(* IEC 61131-3 sources: daoli-st-library/DL_MathData (part 16) *)

(* ---- FC_DL_IntIsPrimeUdint.st ---- *)
(*==============================================================================
 * 组件名称 : FC_DL_IntIsPrimeUdint ｜ 子库 : DL_MathData ｜ v1.0.0 ｜ 2026-11-24
 * 平台     : CODESYS 3.5 / TwinCAT 3 / InoProShop / Machine Expert（纯 IEC，无厂商库）
 * 功能简介 : UDINT 素性判定（试除法）。供伪随机序列、哈希桶数选取、周期分解等调用方。
 *            循环条件写作 nD <= nVal / nD，用除法代替 nD × nD，从根上排除乘法溢出（禁 i*i）。
 * 契约     : 返回 TRUE 表示素数、FALSE 表示合数或 nVal < 2；两者均为合法答案，
 *            bValid := TRUE、bError 保持 FALSE（本件无故障级路径，全为信息级语义）。
 * 依赖     : 无 DL_ 内部依赖（R16 自足实现），无标准库函数调用
 * 错误码   : R297 零码位范式：eErr 恒 0，仅以 bError / bValid 表达
 * 红线自检 : R1 零全局 R2 零%I/%Q R3 纯IEC R4 除零前置（nD ≥ 3 恒定）+ 禁 i*i
 *            R5 双语注释 R6 N/A（无状态机）R7 N/A（无定时器/沿实例）
 *            R10 无类型转换 R11 全声明行分号 R15 标识符零保留字冲突
 * 遗留假设 : nVal < 2（含 0、1）非素数；2 为唯一偶素数，其余偶数短路；
 *            循环天然终止（nD 严格递增、nVal / nD 单调递减），故不设守卫计数；
 *            最坏步数 ⌊√(2³²−1)⌋ / 2 ≈ 32768 次，请在毫秒级任务中避免逐周期调用。
 * 修订历史 : 2026-11-24 R79-B 首版（整数数论族 8/8）
 *============================================================================*)
FUNCTION FC_DL_IntIsPrimeUdint : BOOL
VAR_INPUT
    nVal : UDINT := 0; // 待判定整数 [无量纲] / the value to be tested
END_VAR
VAR_OUTPUT
    eErr   : UDINT; // 错误码，零码位范式恒 0 / error id, always zero under the zero-code rule
    bError : BOOL;  // 故障标志，本件恒 FALSE（素性判定无故障级）/ the fault flag, always FALSE here
    bValid : BOOL;  // 返回值可用标志 / TRUE when the return value is usable
END_VAR
VAR CONSTANT
    DL_ZERO  : UDINT := 0; // 无符号零哨兵 / unsigned zero sentinel
    DL_ONE   : UDINT := 1; // 无符号一哨兵 / unsigned one sentinel
    DL_TWO   : UDINT := 2; // 无符号二哨兵，唯一偶素数 / unsigned two, the only even prime
    DL_THREE : UDINT := 3; // 无符号三哨兵，试除起点 / unsigned three, the trial division start
END_VAR
VAR
    nD : UDINT; // 试除因子，仅取奇数 3, 5, 7, … [无量纲] / the odd trial divisor
END_VAR

// 段 1｜出口预置 / segment 1, preset the exit
FC_DL_IntIsPrimeUdint := FALSE;  // 缺省合数 / default to composite
eErr   := 0;                     // 零码位范式 / zero-code rule
bError := FALSE;                 // 本件无故障级 / this component has no fault level
bValid := FALSE;                 // 判定完成前不认出参 / the result is unusable until the decision is made

// 段 2｜小于 2 的域闸：0 与 1 都不是素数，属合法答案不算故障 / segment 2, the lower domain gate
IF nVal < DL_TWO THEN
    bValid := TRUE;              // FALSE 是合法答案 / FALSE is a legal answer
    RETURN;                      // 返回 FALSE / return the preset FALSE
END_IF

// 段 3｜2 与偶数短路：2 是唯一偶素数 / segment 3, the two and the even number short circuits
IF nVal = DL_TWO THEN
    FC_DL_IntIsPrimeUdint := TRUE;  // 2 为素数 / two is prime
    bValid := TRUE;                 // 判定可用 / the decision is usable
    RETURN;                         // 返回 TRUE / return TRUE
END_IF
IF (nVal MOD DL_TWO) = DL_ZERO THEN
    bValid := TRUE;              // 合数是合法答案 / composite is a legal answer
    RETURN;                      // 返回 FALSE / return the preset FALSE
END_IF

// 段 4｜奇数试除：条件写 nD <= nVal / nD，等价于 nD² <= nVal 但永不溢出 / segment 4, the odd trial division
nD := DL_THREE;                  // 试除起点 3 / start from three
WHILE nD <= (nVal / nD) DO       // 除零不可达：nD ≥ 3 / the divisor is at least three, so no division by zero
    IF (nVal MOD nD) = DL_ZERO THEN
        bValid := TRUE;          // 合数是合法答案 / composite is a legal answer
        RETURN;                  // 返回 FALSE / return the preset FALSE
    END_IF
    nD := nD + DL_TWO;           // 只试奇数 / odd divisors only
END_WHILE

// 段 5｜无因子即素数 / segment 5, no divisor means prime
FC_DL_IntIsPrimeUdint := TRUE;   // 素数 / prime
bValid := TRUE;                  // 判定可用 / the decision is usable
END_FUNCTION

(* ---- FC_DL_IntLcmSafeUdint.st ---- *)
(*==============================================================================
 * 组件名称 : FC_DL_IntLcmSafeUdint ｜ 子库 : DL_MathData ｜ v1.0.0 ｜ 2026-11-24
 * 平台     : CODESYS 3.5 / TwinCAT 3 / InoProShop / Machine Expert（纯 IEC，无厂商库）
 * 功能简介 : UDINT 最小公倍数，先除后乘防溢出：LCM = (nA / GCD) × nB。供脉冲当量配比、
 *            电子齿轮比约分、多轴同步周期归一使用。
 * 契约     : 任一入参为 0 返回 0（IV 约定 LCM(0, x) = 0，信息级，bError 保持 FALSE）；
 *            乘积仍溢出 UDINT 时饱和到 16#FFFF_FFFF 并置 bOverflow := TRUE、bError := TRUE、
 *            bValid := FALSE（饱和值非精确结果，调用方须按故障处理）。
 * 依赖     : 无 DL_ 内部依赖（R16 自足实现：欧几里得 GCD 内联），无标准库函数调用
 * 错误码   : R297 零码位范式：eErr 恒 0，仅以 bError / bValid / bOverflow 表达
 * 红线自检 : R1 零全局 R2 零%I/%Q R3 纯IEC R4 除零前置（nG ≥ 1 由「非双零」保证）+ 乘法前反算上界
 *            R5 双语注释 R6 N/A（无状态机）R7 N/A（无定时器/沿实例）
 *            R10 无类型转换 R11 全声明行分号 R15 标识符零保留字冲突
 * 遗留假设 : 双零入参同属「任一为 0」分支返回 0；GCD 迭代守卫 64 步为安全断言，
 *            理论不可达（欧几里得余量单调递减）；溢出判定用 nQ > (16#FFFF_FFFF / nB)
 *            反算，不做乘法后再比（乘后比已无意义，值已回绕）。
 * 修订历史 : 2026-11-24 R79-B 首版（整数数论族 7/8）
 *============================================================================*)
FUNCTION FC_DL_IntLcmSafeUdint : UDINT
VAR_INPUT
    nA : UDINT := 0; // 左操作数 [脉冲 / 计数] / the left operand, unsigned
    nB : UDINT := 0; // 右操作数 [脉冲 / 计数] / the right operand, unsigned
END_VAR
VAR_OUTPUT
    eErr      : UDINT; // 错误码，零码位范式恒 0 / error id, always zero under the zero-code rule
    bError    : BOOL;  // 乘积溢出时为真（与 bOverflow 同源）/ TRUE on a product overflow, the same source as bOverflow
    bValid    : BOOL;  // 返回值可用标志 / TRUE when the return value is usable
    bOverflow : BOOL;  // 饱和标志：已钳到 16#FFFF_FFFF / TRUE when the result is saturated to the unsigned ceiling
END_VAR
VAR CONSTANT
    DL_ZERO  : UDINT := 0;          // 无符号零哨兵 / unsigned zero sentinel
    DL_ONE   : UDINT := 1;          // 无符号一哨兵 / unsigned one sentinel
    DL_UMAX  : UDINT := 16#FFFF_FFFF; // UDINT 上界，饱和目标 [无量纲] / the unsigned ceiling used for saturation
    DL_GUARD : DINT  := 64;         // GCD 迭代守卫上界 [次] / the euclid guard ceiling
    DL_GUARDI : DINT := 0;          // 迭代计数初值 [次] / the iteration counter start value
END_VAR
VAR
    nX    : UDINT; // GCD 迭代被除数副本 [无量纲] / the gcd dividend copy
    nY    : UDINT; // GCD 迭代除数副本 [无量纲] / the gcd divisor copy
    nG    : UDINT; // 最大公约数 [无量纲] / the greatest common divisor
    nQ    : UDINT; // 先除得商 nA / GCD [无量纲] / the quotient of the division done first
    nIter : DINT;  // GCD 迭代计数，供收敛审计 [次] / the euclid iteration count
END_VAR

// 段 1｜出口预置 / segment 1, preset the exit
FC_DL_IntLcmSafeUdint := DL_ZERO;  // 缺省零 / default zero
eErr      := 0;                    // 零码位范式 / zero-code rule
bError    := FALSE;                // 预置无故障 / preset no fault
bValid    := FALSE;                // 域闸前不认返回值 / the return value is unusable until the gates pass
bOverflow := FALSE;                // 预置未饱和 / preset no saturation

// 段 2｜零入参短路：IV 约定 LCM(0, x) = 0，属信息级不算故障 / segment 2, the zero operand short circuit
IF (nA = DL_ZERO) OR (nB = DL_ZERO) THEN
    bValid := TRUE;                // 0 是合法约定值 / zero is the agreed value here
    RETURN;                        // 返回 0 / return the preset zero
END_IF

// 段 3｜欧几里得 GCD（守卫计数为安全断言，理论不可达）/ segment 3, the euclidean gcd with a guard
nX    := nA;                       // 被除数副本 / dividend copy
nY    := nB;                       // 除数副本 / divisor copy
nIter := DL_GUARDI;                // 计数清零 / clear the counter
WHILE (nY <> DL_ZERO) AND (nIter < DL_GUARD) DO
    nG    := nX MOD nY;            // 余数（nY 非零已证，除法安全）/ the remainder, the divisor is proven non zero
    nX    := nY;                   // 左移 / shift left
    nY    := nG;                   // 左移 / shift left
    nIter := nIter + 1;            // 计数递增 / increment the counter
END_WHILE
IF nIter >= DL_GUARD THEN
    bError := TRUE;                // 守卫命中属平台异常 / a guard hit means a platform anomaly
    RETURN;                        // 返回 0 / return the preset zero
END_IF
nG := nX;                          // 收敛值即 GCD，非双零保证 nG ≥ 1 / the converged value is the gcd and it is at least one

// 段 4｜先除：nQ = nA / GCD，除零已被 nG ≥ 1 拦住 / segment 4, the division done before the multiplication
nQ := nA / nG;                     // 商 [无量纲] / the quotient

// 段 5｜乘法前反算上界：nQ × nB 是否可表示 / segment 5, the pre multiplication ceiling
IF nQ > (DL_UMAX / nB) THEN        // 除零不可达：nB 非零已由段 2 保证 / the divisor is proven non zero
    bOverflow := TRUE;             // 饱和标志 / saturation flag
    bError    := TRUE;             // 故障级：结果不精确 / fault level, the result is inexact
    FC_DL_IntLcmSafeUdint := DL_UMAX;  // 饱和到上界 / saturate to the ceiling
    RETURN;                        // bValid 保持 FALSE / bValid stays FALSE
END_IF

// 段 6｜安全乘法与出口 / segment 6, the safe multiplication and the exit
FC_DL_IntLcmSafeUdint := nQ * nB;  // 已证可表示 / proven representable
bValid := TRUE;                    // 返回值可用 / the return value is usable
END_FUNCTION

(* ---- FC_DL_IntModChk.st ---- *)
(*
    FC_DL_IntModChk —— DINT 整数取模防御包装
    ------------------------------------------------------------------
    组件名称  : FC_DL_IntModChk
    分类      : DL_MathData / IntegerMod
    前缀      : FC_DL_
    版本      : 1.0.0
    溯源      : IEC 61131-3 标准语义的道莅防御性实现（IEC 61131-3 第三版
                整数除法「截断向零」条款 + 余数恒等式 r = a − trunc(a/b)·b
                的防御性落地）；取模语义与判据顺序参照库内 LREAL 域属主
                FC_DL_ModLrealSafe 的闸序（库内复用口径），实现 / 引脚名 /
                码位 100% 自有；clean-room 声明 —— 零代码行复制，无闭源参考。
    平台      : 纯 IEC 61131-3（LINT 64 位整数 + 标准 MOD / DIV 运算符），
                CODESYS 3.5 / TwinCAT 3 / InoProShop / Machine Expert 通用
    作者      : 道莅代码库 · PLC编程专家（R72 构建轮 · 批 1 · 序号 1）
    ------------------------------------------------------------------
    功能说明  : DINT 整数取模 a MOD b 的防御包装，真实工况：齿轮比约分、
                卷绕圈数余量、分度索引回绕前的余数预判。
                判据链顺序：
                ① 除零闸（b = 0 → 故障级早退，输出 0）——先判后除（红线 2）；
                ② DINT_MIN / −1 溢出面闸：被除数 = −2147483648 且除数 = −1 时
                   商 = +2147483648 超出 DINT 可表域（数学余数恒为 0，但三平台
                   MOD 内部实现可能经「先除后乘」路径内溢），此组合显式拦截出
                   信息级，输出确定值 0（数学事实不受影响）；
                ③ 负操作数语义写死：本件**不直接使用平台 MOD 运算符出结果**，
                   而是把两操作数升位到 LINT（64 位，全 DINT 域无损），按
                   IEC 61131-3「整数除法截断向零」标准条款以
                   r = a − trunc(a / b) × b 恒等式自算余数——结果符号**随被除数**
                   （与 C 系 % 口径一致，IEC MOD 主流口径），绝不依赖平台默认；
                ④ 出口（LINT_TO_DINT 降位前已证 |r| < |b| ≤ 2147483648 且
                   r ≠ −2147483648，降位无回绕面）。
                升位理由（可表性反算，R63 口径）：DINT_MIN 取绝对值会在 DINT
                域内回绕（|−2147483648| = 2147483648 > DINT_MAX），任何在
                DINT 域内自算绝对值的写法都带隐藏回绕面；LINT 域内
                ±2147483648 完全可表，升位后全部中间量无回绕。
    错误码    : 16#0002_3900 除数为 0（除零闸命中，输出 0）—— 故障级
                16#0002_3901 被除数 = DINT_MIN 且除数 = −1 的溢出面组合，
                            数学余数恒 0，输出确定值 0、bValid = TRUE —— 信息级，
                            不置 bError（R45）
                加码反证句（R90）：3901 场景（DINT_MIN/−1 组合）无法由「除零码 +
                正常返回值」组合观测——除零码下输出同为 0 但 bValid = FALSE 且
                语义是「除不了」，3901 语义是「可除但实现面危险」，输出组合不可
                互换观测，故立独立码。
    码位总账  : 16#0002_3900 用 ｜ 16#0002_3901 用
    状态机    : N/A —— 纯函数无状态，无 CASE 可写，非法状态不可能出现
    边界与披露: 一 无定时器 / 无沿检测实例 / 无数组下标，周期安全规则 N/A；
                二 零全局变量、零 VAR_EXTERNAL、零物理地址；
                三 整数进位点（终审两式 #2）验收向量：「除子恰为 0」→ 3900
                   故障级输出 0；「被除数 = DINT_MIN 且除子 = −1」→ 3901
                   信息级输出 0；负操作数四象限向量见验收段；
                四 除法面唯一（LINT 域 trunc(a/b)），除数已在段 3 闸为非零，
                   先判后除，无裸除法暴露；
                五 与 FC_DL_ModLrealSafe（DL_MathData，LREAL 浮点域）分工互引：
                   本件只做 DINT 整数域（DINT_MIN/−1 溢出面为浮点域不存在的
                   独立语义），浮点取模一律走属主件，本件不接 LREAL；
                六 依赖声明：仅 Standard.library（无内建函数依赖，LINT 运算符
                   与 DINT_TO_LINT / LINT_TO_DINT 标准转换），三平台无编译门槛。
    验收向量  : V1 (17, 5) → 2；V2 (−17, 5) → −2（符号随被除数）；
                V3 (17, −5) → 2；V4 (−17, −5) → −2；
                V5 (−2147483648, 5) → −3；V6 (−2147483648, −1) → 0 + 3901；
                V7 (x, 0) → 0 + 3900 故障级；V8 (0, 7) → 0。
                算法已证（脚本）：未跑 ｜ 编译器已证（三平台）：未跑
    修订记录  : 2026-11-23 v1.0.0 首次入库（R72 构建轮 · 批 1 · 序号 1）
*)
FUNCTION FC_DL_IntModChk : DINT
VAR_INPUT
    nDividend : DINT;                      (* 被除数，[无量纲整数域] / the dividend, dimensionless integer *)
    nDivisor  : DINT;                      (* 除数，[无量纲整数域]，禁 0 / the divisor, must not be zero *)
END_VAR
VAR_OUTPUT
    bValid    : BOOL;                      (* 返回值（余数）可用标志，故障级为 FALSE / the remainder usable flag, FALSE on fault *)
    bError    : BOOL;                      (* 故障标志，仅故障级码置位（R45 配对）/ the fault flag, raised only on fault level codes *)
    nInfoCode : UDINT;                     (* 信息 / 错误码，0 = 正常 / the info or error id, 0 = ok *)
END_VAR
VAR CONSTANT
    DL_IMD_ZERO   : DINT := 0;             (* 整数零哨兵，除零闸用 [无量纲] / the integer zero sentinel for the divide gate *)
    DL_IMD_DMIN   : DINT := -2147483648;   (* DINT 下界常量（-2^31），溢出面闸用 [无量纲] / the DINT lower bound constant for the overflow gate *)
    DL_IMD_MONE   : DINT := -1;            (* 溢出面除数哨兵 −1 [无量纲] / the overflow gate divisor sentinel *)
END_VAR
VAR
    nLA      : LINT;                       (* 升位被除数（全 DINT 域无损）[无量纲] / the widened dividend *)
    nLB      : LINT;                       (* 升位除数 [无量纲] / the widened divisor *)
    nLQ      : LINT;                       (* LINT 域截断向零商（中间量）[无量纲] / the widened truncating quotient *)
    nLR      : LINT;                       (* LINT 域余数恒等式结果 [无量纲] / the widened remainder *)
END_VAR

// 段 1｜返回值与状态预置（统一出口预置，R256）/ segment 1, preset the return and the status
FC_DL_IntModChk := 0;                      // 故障缺省返回零余数 / the fault default is zero remainder
bValid    := FALSE;                        // 预置不可用，过闸后置位 / preset unusable, set TRUE after the gates
bError    := FALSE;                        // 预置无故障 / preset no fault
nInfoCode := 0;                            // 预置无错 / preset no error
nLA := 0;                                  // 升位中间量清零 / clear the widened dividend
nLB := 0;                                  // 升位中间量清零 / clear the widened divisor
nLQ := 0;                                  // 商中间量清零 / clear the quotient temporary
nLR := 0;                                  // 余数中间量清零 / clear the remainder temporary

// 段 2｜除零闸（先判后除，红线 2；除子恰为 0 验收向量在此命中）/ segment 2, the divide by zero gate
IF nDivisor = DL_IMD_ZERO THEN             // 除数为 0，取模无定义 / the divisor is zero, modulo undefined
    nInfoCode := 16#0002_3900;             // 故障级：除零 / fault level: divide by zero
    bError := TRUE;                        // R45 配对置故障标志 / paired with the fault flag
    bValid := FALSE;                       // 返回值不可用 / the return unusable
    FC_DL_IntModChk := 0;                  // 确定值零出口 / a deterministic zero outlet
    RETURN;                                // 结构早退 / structural exit
END_IF

// 段 3｜DINT_MIN / −1 溢出面闸（商 +2147483648 超 DINT 可表域，防御性拦截）/ segment 3, the DINT_MIN over minus one overflow gate
IF (nDividend = DL_IMD_DMIN) AND (nDivisor = DL_IMD_MONE) THEN // 溢出面组合 / the overflow surface pair
    nInfoCode := 16#0002_3901;             // 信息级：溢出面组合拦截（数学余数恒 0）/ info level: the overflow pair intercepted, the remainder is zero
    bError := FALSE;                       // 信息级不置故障（R45 配对纪律）/ info level never raises a fault
    bValid := TRUE;                        // 数学余数恒为 0，值可用 / the mathematical remainder is zero, usable
    FC_DL_IntModChk := 0;                  // 确定值零出口 / a deterministic zero outlet
    RETURN;                                // 结构早退 / exit
END_IF

// 段 4｜升位与余数恒等式（负操作数语义写死：r = a − trunc(a/b)·b，符号随被除数）/ segment 4, widen and apply the remainder identity
nLA := DINT_TO_LINT(nDividend);            // 被除数升位（全 DINT 域无损）/ widen the dividend lossless
nLB := DINT_TO_LINT(nDivisor);             // 除数升位 / widen the divisor
nLQ := nLA / nLB;                          // IEC 整数除法截断向零（除数已过闸非零）/ the IEC truncating division, divisor gated non zero
nLR := nLA - (nLQ * nLB);                  // 余数恒等式（符号随被除数，不依赖平台 MOD 口径）/ the remainder identity, sign follows the dividend

// 段 5｜降位可表性防线（|r| < |b| ≤ 2147483648 且 r ≠ −2147483648，结构性可证）/ segment 5, the narrowing guard
IF (nLR > DINT_TO_LINT(2147483647)) OR (nLR < DINT_TO_LINT(DL_IMD_DMIN)) THEN // 降位越域防御兜底（不可达，R151 收口纪律）/ the narrowing overflow guard, structurally unreachable
    nInfoCode := 16#0002_3900;             // 复用除零故障级（同属「结果不可信」类，R90 反证：不可达无观测需求）/ reuse the fault code, unreachable
    bError := TRUE;                        // R45 配对置故障标志 / paired with the fault flag
    bValid := FALSE;                       // 返回值不可用 / unusable
    FC_DL_IntModChk := 0;                  // 确定值零出口 / a deterministic zero outlet
    RETURN;                                // 结构早退 / exit
END_IF

// 段 6｜正常出口 / segment 6, the normal outlet
FC_DL_IntModChk := LINT_TO_DINT(nLR);      // 降位发布余数（符号随被除数）/ publish the remainder
bValid := TRUE;                            // 结果可用 / the result usable
END_FUNCTION

(* ---- FC_DL_IntModPowUdint.st ---- *)
(*==============================================================================
 * 组件名称 : FC_DL_IntModPowUdint ｜ 子库 : DL_MathData ｜ v1.0.0 ｜ 2026-11-24
 * 平台     : CODESYS 3.5 / TwinCAT 3 / InoProShop / Machine Expert（纯 IEC，无厂商库）
 * 功能简介 : 模幂运算，返回 nBase^nExp MOD nMod。供校验码、伪随机、整数密钥类运算调用方。
 *            防乘溢出：任何一次乘法都拆成 32 步「加倍-加法」，每步先以「nMod − 加数 是否
 *            够减」判进位再即时归约，故累加积与倍增被乘数恒 < nMod，全程不出现回绕。
 * 契约     : nMod = 0 → 返回 0、bError := TRUE（模数缺失，模幂无定义）；
 *            nMod = 1 → 返回 0、bValid := TRUE（任何数模 1 恒 0，非故障）；
 *            其余 → 返回精确结果、bValid := TRUE、bError 保持 FALSE。
 * 依赖     : 无 DL_ 内部依赖（R16 自足实现：快速乘内联），无标准库函数调用
 * 错误码   : R297 零码位范式：eErr 恒 0，仅以 bError / bValid 表达
 * 红线自检 : R1 零全局 R2 零%I/%Q R3 纯IEC R4 除零前置（nMod ≥ 2 后才有 MOD 与除）+ 乘前归约
 *            R5 双语注释 R6 N/A（无状态机）R7 N/A（无定时器/沿实例）
 *            R10 无类型转换 R11 全声明行分号 R15 标识符零保留字冲突
 * 遗留假设 : 指数位宽固定 UDINT 32 位（内层 FOR 0..31 定长）；两路乘法（nRes × nPow 与
 *            nPow × nPow）合并进同一 32 步循环并行累加，指数位为 0 时积 1 算出后丢弃
 *            （换来「一段代码两用、零重复」，代价是每外层位最多 32 步空转）；
 *            末位之后多做一次倍增无害（nDbl 恒 < nMod），故不设位序守卫。
 * 修订历史 : 2026-11-24 R79-B 首版（整数数论族 9/8 补位）
 *============================================================================*)
FUNCTION FC_DL_IntModPowUdint : UDINT
VAR_INPUT
    nBase : UDINT := 0; // 底数 [无量纲] / the base of the power
    nExp  : UDINT := 0; // 指数 [无量纲] / the exponent
    nMod  : UDINT := 0; // 模数，须 ≥ 2 才有意义 [无量纲] / the modulus, meaningful from two upwards
END_VAR
VAR_OUTPUT
    eErr   : UDINT; // 错误码，零码位范式恒 0 / error id, always zero under the zero-code rule
    bError : BOOL;  // 模数为零时为真 / TRUE when the modulus is zero
    bValid : BOOL;  // 返回值可用标志 / TRUE when the return value is usable
END_VAR
VAR CONSTANT
    DL_ZERO : UDINT := 0; // 无符号零哨兵 / unsigned zero sentinel
    DL_ONE  : UDINT := 1; // 无符号一哨兵 / unsigned one sentinel
    DL_TWO  : UDINT := 2; // 无符号二哨兵，右移与奇偶判据 / unsigned two, the halving and parity base
    DL_BIT0 : DINT  := 0;  // 位循环起点 [位] / the bit loop start index
    DL_BITN : DINT  := 31; // 位循环终点，UDINT 位宽减一 [位] / the bit loop end index
END_VAR
VAR
    nRes  : UDINT; // 结果累加量，恒 < nMod [无量纲] / the result accumulator, always below the modulus
    nPow  : UDINT; // 当前幂底，恒 < nMod [无量纲] / the current power base, always below the modulus
    nExpW : UDINT; // 指数工作副本，逐位右移 [无量纲] / the exponent working copy, shifted per bit
    nMr   : UDINT; // 乘法 1 的乘数（结果量）[无量纲] / the multiplier of the first product
    nMq   : UDINT; // 乘法 2 的乘数（幂底自乘）[无量纲] / the multiplier of the squaring product
    nDbl  : UDINT; // 共用的倍增被乘数，恒 < nMod [无量纲] / the shared doubled multiplicand, always below the modulus
    nAdd  : UDINT; // 本步实际加数，位为 0 时取 0 [无量纲] / the addend of this step, zero on a cleared bit
    nAccR : UDINT; // 乘法 1 的积，恒 < nMod [无量纲] / the accumulator of the first product
    nAccQ : UDINT; // 乘法 2 的积，恒 < nMod [无量纲] / the accumulator of the squaring product
    nBit  : DINT;  // 位循环计数 0..31 [位] / the bit loop counter
END_VAR

// 段 1｜出口预置 / segment 1, preset the exit
FC_DL_IntModPowUdint := DL_ZERO;  // 缺省零 / default zero
eErr   := 0;                      // 零码位范式 / zero-code rule
bError := FALSE;                  // 预置无故障 / preset no fault
bValid := FALSE;                  // 域闸前不认返回值 / the return value is unusable until the gates pass

// 段 2｜模数域闸：零模数故障、一模数恒零 / segment 2, the modulus gates
IF nMod = DL_ZERO THEN
    bError := TRUE;               // 模数缺失，模幂无定义 / without a modulus the operation is undefined
    RETURN;                       // 返回 0 / return the preset zero
END_IF
IF nMod = DL_ONE THEN
    bValid := TRUE;               // 任何数模 1 恒 0，属合法结果 / any value modulo one is zero, a legal result
    RETURN;                       // 返回 0 / return the preset zero
END_IF

// 段 3｜初值：nRes = 1、nPow = nBase MOD nMod（nMod ≥ 2 已证，MOD 安全）/ segment 3, the initial values
nRes  := DL_ONE;                  // 乘法单位元 / the multiplicative identity
nPow  := nBase MOD nMod;          // 底数先归约 / reduce the base first
nExpW := nExp;                    // 指数工作副本 / the exponent working copy

// 段 4｜二进制模幂：指数位自低向高，每轮并行算 nRes × nPow 与 nPow × nPow / segment 4, the binary modular power
WHILE nExpW > DL_ZERO DO
    nMr   := nRes;                // 乘法 1 的乘数 / the first multiplier
    nMq   := nPow;                // 乘法 2 的乘数 / the squaring multiplier
    nDbl  := nPow;                // 两路共用被乘数 / the shared multiplicand
    nAccR := DL_ZERO;             // 积 1 清零 / clear the first accumulator
    nAccQ := DL_ZERO;             // 积 2 清零 / clear the second accumulator
    FOR nBit := DL_BIT0 TO DL_BITN DO
        nAdd := DL_ZERO;                                                     // 加数缺省 0（位为 0 即空加）/ default addend, an empty add on a cleared bit
        IF (nMr MOD DL_TWO) = DL_ONE THEN nAdd := nDbl; END_IF               // 位为 1 才置加数 / load the addend on a set bit
        IF nAccR >= (nMod - nAdd) THEN nAccR := nAccR - (nMod - nAdd); ELSE nAccR := nAccR + nAdd; END_IF  // 加后即时归约，永不溢出 / add and reduce at once
        nAdd := DL_ZERO;                                                     // 加数复用前清零 / clear the reused addend
        IF (nMq MOD DL_TWO) = DL_ONE THEN nAdd := nDbl; END_IF               // 平方路的同款取数 / the same pick for the squaring
        IF nAccQ >= (nMod - nAdd) THEN nAccQ := nAccQ - (nMod - nAdd); ELSE nAccQ := nAccQ + nAdd; END_IF  // 平方路累加 / accumulate the squaring
        nMr := nMr / DL_TWO;                                                 // 乘数 1 右移一位 / shift the first multiplier
        nMq := nMq / DL_TWO;                                                 // 乘数 2 右移一位 / shift the second multiplier
        IF nDbl >= (nMod - nDbl) THEN nDbl := nDbl - (nMod - nDbl); ELSE nDbl := nDbl + nDbl; END_IF        // 被乘数倍增 mod nMod / double the multiplicand modulo the modulus
    END_FOR
    IF (nExpW MOD DL_TWO) = DL_ONE THEN nRes := nAccR; END_IF                // 指数位为 1 才采信积 1 / adopt the first product only on a set exponent bit
    nPow  := nAccQ;               // 平方结果无条件生效 / the squaring always takes effect
    nExpW := nExpW / DL_TWO;      // 指数右移一位 / shift the exponent
END_WHILE

// 段 5｜出口 / segment 5, the exit
FC_DL_IntModPowUdint := nRes;     // 回写结果 / publish the result
bValid := TRUE;                   // 返回值可用 / the return value is usable
END_FUNCTION

(* ---- FC_DL_IntNextPrimeUdint.st ---- *)
(*==============================================================================
 * 组件名称 : FC_DL_IntNextPrimeUdint ｜ 子库 : DL_MathData ｜ v1.0.0 ｜ 2026-11-24
 * 平台     : CODESYS 3.5 / TwinCAT 3 / InoProShop / Machine Expert（纯 IEC，无厂商库）
 * 功能简介 : 求「≥ nVal + 1 的最小素数」（严格大于入参）。供哈希桶数取素数、抖动模数
 *            选取、伪随机种子上限归整使用。试除条件写作 nD <= nCand / nD，禁 i*i 防溢出。
 * 契约     : 找到即返回该素数、bValid := TRUE；nVal ≥ 16#FFFF_FFF0（无足够向上空间）
 *            或 2000 步内未找到（防死循环）或推进中将越过 UDINT 上界 → 返回 0、
 *            bError := TRUE、bValid := FALSE。
 * 依赖     : 无 DL_ 内部依赖（R16 自足实现：试除内联），无标准库函数调用
 * 错误码   : R297 零码位范式：eErr 恒 0，仅以 bError / bValid 表达
 * 红线自检 : R1 零全局 R2 零%I/%Q R3 纯IEC R4 除零前置（nD ≥ 2）+ 步数上限 + 加法溢出兜底
 *            R5 双语注释 R6 N/A（无状态机）R7 N/A（无定时器/沿实例）
 *            R10 无类型转换 R11 全声明行分号 R15 标识符零保留字冲突
 * 遗留假设 : nVal = 0 或 1 时起点取 2（2 是 ≥ 2 的最小素数）；候选逐 1 递增（不跳偶），
 *            保证 2000 步覆盖 2000 个连续整数，远大于 2³² 内的最大素数间隙（≈336），
 *            故「步数命中」只可能发生在接近上界处，与上界兜底互为双保险。
 * 修订历史 : 2026-11-24 R79-B 首版（整数数论族补位）
 *============================================================================*)
FUNCTION FC_DL_IntNextPrimeUdint : UDINT
VAR_INPUT
    nVal : UDINT := 0; // 参考值，本件返回严格大于它的最小素数 [无量纲] / the reference value, the result is strictly above it
END_VAR
VAR_OUTPUT
    eErr   : UDINT; // 错误码，零码位范式恒 0 / error id, always zero under the zero-code rule
    bError : BOOL;  // 无解或搜索步数越界时为真 / TRUE when no answer exists or the search budget is exhausted
    bValid : BOOL;  // 返回值可用标志 / TRUE when the return value is usable
END_VAR
VAR CONSTANT
    DL_ZERO  : UDINT := 0;            // 无符号零哨兵 / unsigned zero sentinel
    DL_ONE   : UDINT := 1;            // 无符号一哨兵 / unsigned one sentinel
    DL_TWO   : UDINT := 2;            // 无符号二哨兵，最小素数 / unsigned two, the smallest prime
    DL_THREE : UDINT := 3;            // 无符号三哨兵，试除起点 / unsigned three, the trial division start
    DL_NEAR  : UDINT := 16#FFFF_FFF0; // 上界保护带起点，超过即判无解 / the guard band start near the ceiling
    DL_GUARD : UDINT := 16#FFFF_FFFE; // 推进溢出兜底线 / the increment overflow guard line
    DL_STEP  : DINT  := 2000;         // 候选搜索步数预算 [步] / the candidate search budget
    DL_STEP0 : DINT  := 0;            // 步数计数初值 [步] / the step counter start value
    DL_STEP1 : DINT  := 1;            // 步数计数步长 [步] / the step counter increment
END_VAR
VAR
    nCand  : UDINT; // 当前候选整数 [无量纲] / the current candidate
    nD     : UDINT; // 试除因子，奇数 3, 5, 7, … [无量纲] / the odd trial divisor
    nStep  : DINT;  // 已消耗的候选步数 [步] / the consumed candidate steps
    bPrime : BOOL;  // 当前候选的素性结论 / the primality verdict of the current candidate
    bFound : BOOL;  // 找到标志 / the found flag
END_VAR

// 段 1｜出口预置 / segment 1, preset the exit
FC_DL_IntNextPrimeUdint := DL_ZERO;  // 缺省零哨兵 / default zero sentinel
eErr    := 0;                        // 零码位范式 / zero-code rule
bError  := FALSE;                    // 预置无故障 / preset no fault
bValid  := FALSE;                    // 域闸前不认返回值 / the return value is unusable until the gates pass

// 段 2｜上界域闸：无足够向上空间即判无解 / segment 2, the ceiling gate
IF nVal >= DL_NEAR THEN
    bError := TRUE;                  // 上界保护带内不搜索 / no search inside the guard band
    RETURN;                          // 返回 0 / return the preset zero
END_IF

// 段 3｜起点：严格大于入参，且不低于 2 / segment 3, the start candidate
nCand  := nVal + DL_ONE;             // 严格大于入参 / strictly above the argument
IF nCand < DL_TWO THEN nCand := DL_TWO; END_IF  // 0/1 的最小数答案是 2 / two is the answer for zero and one
nStep  := DL_STEP0;                  // 步数清零 / clear the step counter
bFound := FALSE;                     // 未找到 / nothing found yet

// 段 4｜候选搜索：逐 1 递增，超出预算即停（防死循环）/ segment 4, the candidate search
WHILE (NOT bFound) AND (nStep < DL_STEP) DO
    nStep  := nStep + DL_STEP1;      // 消耗一步 / consume one step
    bPrime := TRUE;                  // 先假定素数 / assume prime first
    IF (nCand > DL_TWO) AND ((nCand MOD DL_TWO) = DL_ZERO) THEN bPrime := FALSE; END_IF  // 大于 2 的偶数必合数 / every even number above two is composite
    IF bPrime AND (nCand > DL_THREE) THEN
        nD := DL_THREE;              // 试除起点 3 / start from three
        WHILE nD <= (nCand / nD) DO  // 等价于 nD² ≤ nCand 但永不溢出 / equivalent to the square test without overflow
            IF (nCand MOD nD) = DL_ZERO THEN
                bPrime := FALSE;     // 找到因子即合数 / a divisor means composite
                EXIT;                // 跳出试除循环 / leave the trial division loop
            END_IF
            nD := nD + DL_TWO;       // 只试奇数 / odd divisors only
        END_WHILE
    END_IF
    IF bPrime THEN
        bFound := TRUE;              // 候选即答案 / the candidate is the answer
    ELSIF nCand >= DL_GUARD THEN
        bError := TRUE;              // 再推进将越过上界 / another step would overflow the ceiling
        bFound := TRUE;              // 以故障方式结束搜索 / end the search as a fault
        nCand  := DL_ZERO;           // 结果置零哨兵 / force the zero sentinel
    ELSE
        nCand := nCand + DL_ONE;     // 推进到下一候选 / advance to the next candidate
    END_IF
END_WHILE

// 段 5｜出口：未找到（预算耗尽）判故障，找到则回写 / segment 5, the exit
IF (NOT bFound) OR bError THEN
    bError := TRUE;                  // 预算耗尽或无解 / the budget ran out or no answer exists
    RETURN;                          // 返回 0 哨兵 / return the zero sentinel
END_IF
FC_DL_IntNextPrimeUdint := nCand;    // 回写素数 / publish the prime
bValid := TRUE;                      // 返回值可用 / the return value is usable
END_FUNCTION

(* ---- FC_DL_IntPowSatUdint.st ---- *)
(*==============================================================================
 * 组件名称 : FC_DL_IntPowSatUdint ｜ 子库 : DL_MathData ｜ v1.0.2 ｜ 2026-11-24
 * 平台     : CODESYS 3.5 / TwinCAT 3 / InoProShop / Machine Expert（纯 IEC，无厂商库）
 * 功能简介 : 无符号整数快速幂（平方求幂），溢出即饱和到 16#FFFF_FFFF 并置 bOverflow。
 *            乘前反算上界：被乘数 > 上限 DIV 乘数 即判溢出，绝不让乘法先回绕。
 * 契约     : 返回 nBase^nExp；nExp = 0 返回 1（含 0^0 口径取 1）；饱和时返回
 *            16#FFFF_FFFF 且 bOverflow := TRUE，bValid 仍为 TRUE（饱和值是确定结论）。
 * 依赖     : 无 DL_ 内部依赖（R16 自足实现），无标准库函数调用
 * 错误码   : R297 零码位范式：eErr 恒 0，饱和以 bOverflow 表达
 * 红线自检 : R1 零全局 R2 零%I/%Q R3 纯IEC R4 乘前反算防溢出、除零前置、循环上限 32 次
 *            R5 双语注释 R6 N/A（无状态机）R7 N/A（无定时器/沿实例）
 *            R10 无类型转换 R11 全声明行分号 R15 标识符零保留字冲突 R18 N/A（无 bReset）
 * 修订历史 : 2026-11-24 R79-A 首版（整数数论族 5/8）
 *============================================================================*)
FUNCTION FC_DL_IntPowSatUdint : UDINT
VAR_INPUT
    nBase       : UDINT;    // 底数，全域 [无量纲] / base over the whole unsigned range
    nExp        : UDINT;    // 指数，全域 [无量纲] / exponent over the whole unsigned range
END_VAR
VAR_OUTPUT
    eErr        : UDINT;    // 错误码，零码位范式恒 0 / error id, always zero under the zero-code rule
    bError      : BOOL;     // 故障标志，本件结构性不置位 / fault flag, never raised by this component
    bValid      : BOOL;     // 结果可用标志，饱和亦为可用结论 / TRUE even when saturated, saturation is a definite verdict
    bOverflow   : BOOL;     // 结果已饱和到 UDINT 上界 / TRUE when the result saturated at the unsigned upper bound
END_VAR
VAR CONSTANT
    DL_MAX_UDINT : UDINT := 16#FFFF_FFFF;   // UDINT 上界，饱和目标值 [无量纲] / unsigned upper bound and saturation target
    DL_TWO       : UDINT := 2;              // 指数折半基数 [无量纲] / exponent halving radix
    DL_ONE       : UDINT := 1;              // 整数一 / integer one
    DL_ZERO      : UDINT := 0;              // 整数零哨兵 / integer zero sentinel
    DL_ITER_MAX  : UDINT := 32;             // 指数最多 32 位，迭代上限 [次] / an exponent has at most thirty two bits [count]
END_VAR
VAR
    nBaseUse    : UDINT;    // 迭代中的底数（含平方） / running base, includes the squaring steps
    nExpUse     : UDINT;    // 迭代中的指数（逐次折半） / running exponent, halved every step
    nRes        : UDINT;    // 结果累乘器 / result accumulator
    nIter       : UDINT;    // 已用迭代次数 / iterations consumed so far
END_VAR

// 段 1｜出口预置 / segment 1, preset the exit
FC_DL_IntPowSatUdint := 0;      // 缺省 0 / default zero
eErr      := 0;                 // 零码位范式 / zero-code rule
bError    := FALSE;             // 本件不产生故障级 / this component raises no fault
bValid    := TRUE;              // 全定义域给出确定结论 / a definite verdict for the whole domain
bOverflow := FALSE;             // 预置未饱和 / preset unsaturated
nRes      := DL_ONE;            // 累乘器初值 1 / accumulator starts at one

// 段 2｜零指数边界：任何底数的 0 次幂为 1 / segment 2, the zero exponent boundary
IF nExp = DL_ZERO THEN
    FC_DL_IntPowSatUdint := DL_ONE;     // 结果为 1 / the result is one
    RETURN;
END_IF

// 段 3｜平方求幂：逐位判断，乘前反算溢出 / segment 3, square and multiply with an overflow reflection
nBaseUse := nBase;                  // 底数工作副本 / working copy of the base
nExpUse  := nExp;                   // 指数工作副本 / working copy of the exponent
nIter    := DL_ZERO;
WHILE (nExpUse > DL_ZERO) AND (nIter < DL_ITER_MAX) DO
    nIter := nIter + DL_ONE;                        // 守卫自增 / advance the guard
    IF (nExpUse MOD DL_TWO) = DL_ONE THEN           // 当前最低位为 1 才乘 / multiply only when the low bit is set
        IF (nBaseUse <> DL_ZERO) AND (nRes > (DL_MAX_UDINT / nBaseUse)) THEN
            nRes      := DL_MAX_UDINT;              // 反算超界，直接饱和 / the reflection overshoots, saturate at once
            bOverflow := TRUE;
        ELSE
            nRes := nRes * nBaseUse;                // 安全乘法 / safe multiplication
        END_IF
    END_IF
    nExpUse := nExpUse / DL_TWO;                    // 指数折半，除数为常量 2 / halve the exponent
    IF nExpUse > DL_ZERO THEN
        IF (nBaseUse <> DL_ZERO) AND (nBaseUse > (DL_MAX_UDINT / nBaseUse)) THEN
            nBaseUse  := DL_MAX_UDINT;              // 平方超界，钳到上限 / the squaring overshoots, clamp to the ceiling
            bOverflow := TRUE;                      // 平方已越界 = 真溢出（v1.0.2 修：v1.0.1 前此处无回执，静默出残值）/ squaring overflowed, raise the receipt (silent residue before v1.0.2)
        ELSE
            nBaseUse := nBaseUse * nBaseUse;        // 安全平方 / safe squaring
        END_IF
    END_IF
END_WHILE
(* v1.0.2 更正：v1.0.1 曾在此按 nIter 触顶置 bOverflow，但 nBase <= 1 且 nExp >= 2^31 时
   循环合法打满 32 次仍应收敛（1^N = 1），该判据造成假溢出回执，已删除；
   溢出回执改为只在「乘前反算越界」与「平方钳位」两处产生（唯一真溢出来源）。 *)

// 段 4｜出口 / segment 4, exit
FC_DL_IntPowSatUdint := nRes;                   // 结果或饱和值 / the result or the saturation value
END_FUNCTION

(* ---- FC_DL_IntReverseDigitsUdint.st ---- *)
(*==============================================================================
 * 组件名称 : FC_DL_IntReverseDigitsUdint ｜ 子库 : DL_MathData ｜ v1.0.0 ｜ 2026-11-24
 * 平台     : CODESYS 3.5 / TwinCAT 3 / InoProShop / Machine Expert（纯 IEC，无厂商库）
 * 功能简介 : 无符号整数的十进制数字反转（如 123 → 321，120 → 21，末尾零自然丢弃）。
 *            逐位取余乘十再累加，纯整数实现。乘前反算：累加器 > (上界 − 当前位) DIV 10
 *            即判溢出，饱和到 16#FFFF_FFFF 并置 bOverflow。
 * 契约     : 返回反转值；反转结果超 UDINT 域时返回 16#FFFF_FFFF、bOverflow := TRUE、
 *            bValid 保持 TRUE（饱和值是确定结论）。nVal = 0 返回 0。
 * 依赖     : 无 DL_ 内部依赖（R16 自足实现），无标准库函数调用
 * 错误码   : R297 零码位范式：eErr 恒 0，溢出以 bOverflow 表达
 * 红线自检 : R1 零全局 R2 零%I/%Q R3 纯IEC R4 乘前反算防溢出、循环上界 10 次、除数为常量
 *            R5 双语注释 R6 N/A（无状态机）R7 N/A（无定时器/沿实例）
 *            R10 无类型转换 R11 全声明行分号 R15 标识符零保留字冲突 R18 N/A（无 bReset）
 * 修订历史 : 2026-11-24 R79-A 首版（整数数论族 8/8）
 *============================================================================*)
FUNCTION FC_DL_IntReverseDigitsUdint : UDINT
VAR_INPUT
    nVal        : UDINT;    // 待反转整数，全域 0~16#FFFF_FFFF [无量纲] / value to reverse over the whole unsigned range
END_VAR
VAR_OUTPUT
    eErr        : UDINT;    // 错误码，零码位范式恒 0 / error id, always zero under the zero-code rule
    bError      : BOOL;     // 故障标志，本件结构性不置位 / fault flag, never raised by this component
    bValid      : BOOL;     // 结果可用标志，饱和亦为可用结论 / TRUE even when saturated
    bOverflow   : BOOL;     // 反转结果已饱和到 UDINT 上界 / TRUE when the reversed value saturated
END_VAR
VAR CONSTANT
    DL_TEN       : UDINT := 10;             // 十进制基数 [无量纲] / decimal radix, dimensionless
    DL_MAX_UDINT : UDINT := 16#FFFF_FFFF;   // UDINT 上界，饱和目标值 [无量纲] / unsigned upper bound and saturation target
    DL_ZERO      : UDINT := 0;              // 整数零哨兵 / integer zero sentinel
    DL_LOOP_MAX  : UDINT := 10;             // UDINT 十进制最大位数，循环上界 [位] / loop cap equal to the largest decimal width [digit]
END_VAR
VAR
    nRest       : UDINT;    // 降位过程中的剩余值 / remaining value while descending
    nRev        : UDINT;    // 反转累加器 / reversed accumulator
    nDigit      : UDINT;    // 当前取出的个位数 / the digit taken from the current position
    nGuard      : UDINT;    // 循环守卫计数 / loop guard counter
END_VAR

// 段 1｜出口预置 / segment 1, preset the exit
FC_DL_IntReverseDigitsUdint := 0;   // 缺省 0 / default zero
eErr      := 0;                     // 零码位范式 / zero-code rule
bError    := FALSE;                 // 本件不产生故障级 / this component raises no fault
bValid    := TRUE;                  // 饱和也是确定结论 / saturation is still a definite verdict
bOverflow := FALSE;                 // 预置未饱和 / preset unsaturated
nRest     := nVal;                  // 从输入起步 / start from the input
nRev      := DL_ZERO;               // 累加器清零 / clear the accumulator
nGuard    := DL_ZERO;               // 守卫清零 / clear the guard

// 段 2｜逐位反转：取个位 → 降位 → 乘前反算后累加 / segment 2, digit by digit reversal with an overflow reflection
WHILE (nRest <> DL_ZERO) AND (nGuard < DL_LOOP_MAX) DO
    nGuard := nGuard + 1;                                   // 守卫自增 / advance the guard
    nDigit := nRest MOD DL_TEN;                             // 取个位 / take the units digit
    nRest  := nRest / DL_TEN;                               // 降一位 / shift one digit down
    IF nRev > ((DL_MAX_UDINT - nDigit) / DL_TEN) THEN
        nRev      := DL_MAX_UDINT;                          // 反算超界，饱和退出 / the reflection overshoots, saturate and stop
        bOverflow := TRUE;
        EXIT;
    END_IF
    nRev := (nRev * DL_TEN) + nDigit;                       // 旧位左移一位并接上新位 / shift the old digits and append
END_WHILE

// 段 3｜出口 / segment 3, exit
FC_DL_IntReverseDigitsUdint := nRev;    // 反转值或饱和值 / the reversed value or the saturation value
END_FUNCTION

(* ---- FC_DL_IntSqrtFloorUdint.st ---- *)
(*==============================================================================
 * 组件名称 : FC_DL_IntSqrtFloorUdint ｜ 子库 : DL_MathData ｜ v1.0.0 ｜ 2026-11-24
 * 平台     : CODESYS 3.5 / TwinCAT 3 / InoProShop / Machine Expert（纯 IEC，无厂商库）
 * 功能简介 : 无符号整数平方根向下取整 ⌊√nVal⌋。牛顿迭代：初值 nVal DIV 2 + 1，
 *            下一试值 = (试值 + nVal DIV 试值) DIV 2，试值不再下降即收敛。
 *            纯整数运算，无浮点、无 SQRT，2^32 全域精确。
 * 契约     : 返回 ⌊√nVal⌋；nVal = 0 返回 0；nIter 达上限 64 次仍未收敛时返回最后一次
 *            试值并置 bError（结构性不可达，作为防死循环兜底）。
 * 依赖     : 无 DL_ 内部依赖（R16 自足实现），无标准库函数调用
 * 错误码   : R297 零码位范式：eErr 恒 0，仅以 bError / bValid 表达
 * 红线自检 : R1 零全局 R2 零%I/%Q R3 纯IEC R4 除零前置（试值恒 ≥1）、迭代上限兜底、
 *            和式上界 ≤ 2^31+1 不溢出 R5 双语注释 R6 N/A（无状态机）
 *            R7 N/A（无定时器/沿实例）R10 无类型转换 R11 全声明行分号
 *            R15 标识符零保留字冲突 R18 N/A（无 bReset）
 * 修订历史 : 2026-11-24 R79-A 首版（整数数论族 1/8）
 *============================================================================*)
FUNCTION FC_DL_IntSqrtFloorUdint : UDINT
VAR_INPUT
    nVal        : UDINT;    // 被开方数，全域 0~16#FFFF_FFFF [无量纲] / radicand over the whole unsigned range
END_VAR
VAR_OUTPUT
    eErr        : UDINT;    // 错误码，零码位范式恒 0 / error id, always zero under the zero-code rule
    bError      : BOOL;     // 迭代未收敛为真（结构性不可达） / TRUE when the iteration fails to converge, unreachable in theory
    bValid      : BOOL;     // 结果可用标志 / result usable flag
END_VAR
VAR CONSTANT
    DL_TWO      : UDINT := 2;               // 牛顿迭代的除数 2 [无量纲] / Newton divisor, dimensionless
    DL_ONE      : UDINT := 1;               // 整数一 [无量纲] / integer one, dimensionless
    DL_ZERO     : UDINT := 0;               // 整数零哨兵 [无量纲] / integer zero sentinel, dimensionless
    DL_ITER_MAX : UDINT := 64;              // 迭代次数上限，二次收敛下 32 次已足 [次] / iteration cap, quadratic convergence needs far fewer [count]
END_VAR
VAR
    nApprox     : UDINT;    // 当前试值，迭代中单调下降 / current trial value, monotonically decreasing
    nNext       : UDINT;    // 下一试值 / next trial value
    nIter       : UDINT;    // 已用迭代次数 / iterations consumed so far
END_VAR

// 段 1｜出口预置 / segment 1, preset the exit
FC_DL_IntSqrtFloorUdint := 0;   // 缺省 0 / default zero
eErr   := 0;                    // 零码位范式 / zero-code rule
bError := FALSE;                // 预置无故障 / preset no fault
bValid := FALSE;                // 计算完成前不认结果 / unusable until the iteration ends

// 段 2｜零边界：0 的平方根为 0，直接放行，避免初值 1 走迭代 / segment 2, the zero boundary
IF nVal = DL_ZERO THEN
    bValid := TRUE;             // 结果 0 可用 / the zero result is usable
    RETURN;                     // 返回 0 / return zero
END_IF

// 段 3｜牛顿迭代：初值取 nVal DIV 2 + 1，必 ≥ √nVal，故单调下降 / segment 3, Newton iteration from an upper bound
nApprox := (nVal / DL_TWO) + DL_ONE;                // 上界初值，避免 nVal DIV nApprox 除零 / upper bound start, keeps the divisor non zero
nIter   := DL_ZERO;                                 // 迭代计数清零 / clear the counter
WHILE nIter < DL_ITER_MAX DO
    nIter   := nIter + DL_ONE;                      // 先计数后算，保证上限生效 / count first so the cap is honoured
    nNext   := (nApprox + (nVal / nApprox)) / DL_TWO;   // 和式上界约 2^31+1，不溢出 / the sum stays near two to the thirty first, no overflow
    IF nNext >= nApprox THEN
        EXIT;                                       // 试值不再下降即收敛 / the trial stops decreasing, converged
    END_IF
    nApprox := nNext;                               // 继续下降 / keep descending
END_WHILE

// 段 4｜收敛自证：用尽上限仍未收敛按故障处置，返回最后一次试值 / segment 4, convergence self proof
IF nIter >= DL_ITER_MAX THEN
    bError := TRUE;                 // 未收敛（理论不可达）/ not converged, unreachable in theory
    FC_DL_IntSqrtFloorUdint := nApprox;
    RETURN;                         // 返回最后一次试值，bValid 保持 FALSE / return the last trial with bValid still FALSE
END_IF

// 段 5｜出口 / segment 5, exit
FC_DL_IntSqrtFloorUdint := nApprox;     // ⌊√nVal⌋ / floor of the square root
bValid := TRUE;                         // 结果可用 / the result is usable
END_FUNCTION

(* ---- FC_DL_IntToFixedField.st ---- *)
(*==============================================================================
 * 组件名称 (Component)  : FC_DL_IntToFixedField
 * 溯源说明 (Provenance): 道莅 clean-room 防御性实现（IEC 61131-3 纯净实现，闭源文档仅借语义，零代码行）
 * 所属子库 (Sublibrary) : DL_MathData / DataFormat
 * 当前版本 (Version)    : 1.0.0
 * 兼容性   (Platform)   : CODESYS 3.5 / TwinCAT 3 / 汇川 InoProShop / 施耐德
 *                         Machine Expert；纯 IEC 61131-3（第 3 版），仅用
 *                         Standard.library 的 MID / CONCAT / LEN
 * 组件分类 (Category)   : 函数（FUNCTION）· 纯函数 · 整数 → 定宽数值字段
 * 功能一句话 (Summary)  : 把 DINT 整数编码成恰好 uWidth 个字符的定宽字段
 *                         （右对齐，零填充或空格填充，可选强制正号），
 *                         供 MES 流水号与 ASCII 定长报文拼装使用。
 *
 * 本件存在的意义 (Why this unit exists)
 *   库内 FC_DL_StringFixedField 解决「定长串填充与对齐」（内容不定），
 *   FC_DL_DintToStringTrim 解决「数值→文本去空格」（不定宽）。二者之间有一个
 *   真实缺口：数值 → **定宽零填充字段**（00012345）与它的逆运算。
 *   MES 流水号、秤重报文、ASCII 定长十进制域全部落在这一格，缺件则报文层
 *   拼不出列位对齐的数字域。本件与 FC_DL_FixedFieldToInt 构成编码对。
 *
 * 【填充与对齐规则（与 FC_DL_FixedFieldToInt 共用同一段口径原文）】
 *   ① 右对齐：数字永远贴字段右端，填充字符只在左侧。
 *   ② 填充字符由 bZeroPad 决定：TRUE 用 '0'，FALSE 用 ' '。
 *   ③ 符号位占一位：零填充时符号贴最左（-0000042），空格填充时符号紧贴数字
 *      （     -42）——这是 C printf 的 %08d / %8d 口径，两种写法的字段长度
 *      都恰好等于 uWidth，任何时刻不会出现半截字段。
 *   ④ 宽度是契约：不够装就**拒绝编码**，绝不截断成半截数字（截断出来的
 *      「1234」与真实「123456」在报文里无法区分，是账实不符的根因）。
 *
 * 边界安全 (Boundary)
 *   ① uWidth < 1 或 > 20 → 钳到 1 / 20 并置信息 045C（宽度可钳，内容不可钳）；
 *   ② 可用数字位（宽度扣掉符号位）不足以容纳全部数字 → 故障 03A8、拒绝编码、
 *      sField 保持空串、uFieldLen 保持 0；
 *   ③ 整数分解**全程走负域**：nValue = -2147483648 若先取绝对值再取模会回绕，
 *      故负值直接进负域、正值先取反进负域，循环内 nWork 恒 ≤ 0，
 *      `-(nWork MOD 10)` 恒得 0~9（IEC：MOD 结果符号随被除数）；
 *   ④ sField 声明 STRING(20) 与本件宽度上限一致，宽度钳位后总长恒 ≤ 20，
 *      写入不存在隐式截断；出口另做 LEN 复检兜底（防御纵深）。
 * 遗留假设 (Assumption)
 *   MOD 的负余数口径按 IEC 61131-3（结果符号随被除数）与 C 语言一致，
 *   本件依赖该口径实现负域分解；CODESYS / TwinCAT / InoProShop 三平台一致。
 *
 * 错误码    : 16#0001_045C 字段宽度越界已钳位到 1~20——信息级，正常防御
 *             16#0001_045D 预留禁用（信息级，不得挪用）
 *             16#0001_03A8 可用宽度不足以容纳完整数值，拒绝编码（不输出半截数字）——故障级，返回 FALSE
 *             16#0001_03A9 预留禁用（故障级，不得挪用）
 *             16#0001_03AA 预留禁用（故障级，不得挪用）
 * 码位总账  : 16#0001_045C 用 / 16#0001_045D 预留 ｜ 16#0001_03A8 用 / 16#0001_03A9 预留 / 16#0001_03AA 预留
 * 状态机    : N/A —— 纯函数无顺序状态机，无 CASE 可写，非法状态不可能出现
 * 采样约定  : 纯组合函数，无定时器、无内部驻留状态，调用即出结果
 * 依赖说明  : 无 DL_ 内部依赖；仅 Standard.library 的 MID / CONCAT / LEN
 * 验收向量  : V1 12345/宽8/零填 → '00012345'，写 8，TRUE
 *             V2 -42/宽8/空格填 → '     -42'，写 8，TRUE
 *             V3 0/宽4/零填 → '0000'
 *             V4 -2147483648/宽11 → '-2147483648'，写 11（负域分解主向量）
 *             V5 123456/宽4 → FALSE，sField=''，uFieldLen=0，eErr=03A8，bError=TRUE
 *             V6 宽 0 → 钳到 1 且 eErr=045C，bError 保持 FALSE
 *             V7 round-trip：#1 编码 → #2 解析，全 DINT 域逐值回原值
 * 红线自检  : 全局变量声明零使用 / 外部变量访问零使用 / 物理地址零使用 ｜ 纯 IEC 61131-3 ｜ 防除零
 *             （本件无除法）· 浮点无比较 · 循环带 nGuard ｜ 全变量双语同行注释
 *             状态机 N/A ｜ 无定时器实例 ｜ 无魔法数（阈值全部 VAR CONSTANT）
 * 修订历史  : 2026-11-16  v1.0.0  首版入库（R22 · 批 1 · 定宽数值字段族）
 *============================================================================*)

FUNCTION FC_DL_IntToFixedField : BOOL
VAR_INPUT
    nValue      : DINT;                        // 待编码整数，全 DINT 域 / integer to encode, full DINT range
    uWidth      : UINT := 8;                   // 字段宽度 [字符]，范围 1~20 / field width [char], range 1~20
    bZeroPad    : BOOL := TRUE;                // TRUE 零填充 / FALSE 空格填充 / TRUE zero padding, FALSE space padding
    bForceSign  : BOOL := FALSE;               // 正数是否强制 '+' 号 / force '+' sign on positive values
END_VAR
VAR_OUTPUT
    sField      : STRING(20);                  // 编码结果，右对齐 [字符] / encoded field, right aligned [char]
    uFieldLen   : UINT;                        // 实际写入字符数 [字符] / actual written length [char]
    eErr        : UDINT;                       // 错误码，0 表示无错 / error code, 0 means no error
    bError      : BOOL;                        // 故障级标志，仅故障级错误置位 / fault-class flag, set only on fault-level codes
    bValid      : BOOL;                        // 结果可用标志 / result usable flag
END_VAR
VAR
    nWUse       : INT;                         // 生效字段宽度 [字符]，已钳位 1~20 / effective width, clamped to 1~20
    nDigitsAvail: INT;                         // 扣符号位后可用数字位 [字符] / digits available after the sign position
    nDigitCount : INT;                         // 实际数字位个数 [位] / actual digit count
    nPadCount   : INT;                         // 填充字符个数 [字符] / pad character count
    nGuard      : INT;                         // 循环守卫计数器 [次] / loop guard counter
    nWork       : DINT;                        // 负域分解工作值，恒 ≤ 0 [无量纲] / negative-domain working value, always <= 0
    nDigit      : DINT;                        // 当前最低位数字 0~9 [无量纲] / current least significant digit
    bNeg        : BOOL;                        // 输入为负数 / input is negative
    bNeedSign   : BOOL;                        // 本字段是否输出符号字符 / whether a sign character is emitted
    sDigits     : STRING(20);                  // 数字段，高位在前 [ASCII] / digit segment, most significant first
    sPad        : STRING(20);                  // 填充段，贴在数字左侧 [ASCII] / pad segment, left of the digits
    sSign       : STRING(1);                   // 符号段，单字符 [ASCII] / sign segment, single character
    sDigitCh    : STRING(1);                   // 单字符数字，由数字表取出 [ASCII] / single digit character taken from the table
END_VAR
VAR CONSTANT
    DL_FIELD_MAX : UINT := 20;                 // STRING(20) 物理上限 [字符]，禁写成 255 / physical bound of STRING(20), never 255
    DL_W_MIN_U   : UINT := 1;                  // 宽度下限的无符号副本 [字符]，用于 UINT 域比较 / unsigned copy of the width lower bound
    DL_W_MIN     : INT := 1;                   // 宽度下限 [字符] / width lower bound [char]
    DL_W_MAX     : INT := 20;                  // 宽度上限 [字符]，与 DL_FIELD_MAX 同值同义 / width upper bound, same value as DL_FIELD_MAX
    DL_DIGIT_MAX : INT := 10;                  // DINT 十进制最大位数 [位] / maximum decimal digits of DINT
    DL_GUARD_MAX : INT := 12;                  // 分解循环守卫上限 [次]，大于位数即安全 / decomposition loop guard, larger than the digit count
    DL_TEN       : DINT := 10;                 // 十进制基数 [无量纲] / decimal radix
    DL_POS_ONE   : INT := 1;                   // MID 的位置基数与单字符长度 [字符] / MID position base and single-char length
    DL_DIGITS    : STRING(10) := '0123456789'; // 数字字符表，经 MID 按下标取值 [ASCII] / digit table indexed through MID
    DL_PAD_ZERO  : STRING(1) := '0';           // 零填充字符 [字符] / zero pad character
    DL_PAD_SPACE : STRING(1) := ' ';           // 空格填充字符 [字符] / space pad character
    DL_SIGN_PLUS : STRING(1) := '+';           // 正号字符 [字符] / plus sign character
    DL_SIGN_MINUS: STRING(1) := '-';           // 负号字符 [字符] / minus sign character
END_VAR

(*------------------------------------------------------------------------------
 * 段 1｜返回值与输出预置（任何早退路径不留脏值，L1/L9）
 *      Preset the return value and every output so no early exit leaves stale data
 *-----------------------------------------------------------------------------*)
FC_DL_IntToFixedField := FALSE;                // 返回值预置失败，成功路径末段置 TRUE / preset to FALSE, set TRUE only on success
sField      := '';                             // 字段清空，拒绝编码时保持空串 / field cleared, stays empty on refusal
uFieldLen   := 0;                              // 写入字符数预置 0 [字符] / written length preset to zero
eErr        := 16#0000_0000;                   // 错误码预置无错 / error code preset to none
bError      := FALSE;                          // 故障标志预置 FALSE / fault flag preset to FALSE
bValid      := FALSE;                          // 结果可用标志预置 FALSE / usable flag preset to FALSE
nWUse       := DL_W_MIN;                       // 生效宽度预置下限 / effective width preset to the lower bound
nDigitsAvail := 0;                             // 可用数字位预置 0 / available digits preset to zero
nDigitCount := 0;                              // 数字位个数预置 0 / digit count preset to zero
nPadCount   := 0;                              // 填充个数预置 0 / pad count preset to zero
nGuard      := 0;                              // 循环守卫预置 0 / guard preset to zero

(*------------------------------------------------------------------------------
 * 段 2｜宽度闸门（越界只钳位不拒绝：宽度可钳，内容不可钳）
 *      Width gate: clamping the width is safe, clamping the content is not
 *-----------------------------------------------------------------------------*)
IF uWidth < DL_W_MIN_U THEN
    nWUse := DL_W_MIN;                         // 钳到下限 1 / clamped to the lower bound
    eErr  := 16#0001_045C;                     // 信息级：宽度已钳位 / informational: width clamped
ELSIF uWidth > DL_FIELD_MAX THEN
    nWUse := DL_W_MAX;                         // 钳到上限 20 / clamped to the upper bound
    eErr  := 16#0001_045C;                     // 信息级：宽度已钳位 / informational: width clamped
ELSE
    nWUse := UINT_TO_INT(uWidth);              // 域内直通 / passed through inside the domain
END_IF

(*------------------------------------------------------------------------------
 * 段 3｜符号判定与可用数字位（符号位先占，再谈数字装不装得下）
 *      Sign decision and available digit positions
 *-----------------------------------------------------------------------------*)
bNeg      := (nValue < 0);                      // 负值判据，DINT 全域成立 / negative test, valid over the whole DINT range
bNeedSign := bNeg OR bForceSign;                // 负号必需，正号由引脚决定 / minus always needed, plus only if forced
IF bNeedSign AND (nWUse >= (DL_W_MIN + DL_POS_ONE)) THEN
    nDigitsAvail := nWUse - DL_POS_ONE;         // 宽度至少 2 才谈得上符号 + 一位数字 / at least two positions for sign plus one digit
ELSIF bNeedSign THEN
    nDigitsAvail := 0;                         // 宽度 1 且要符号：无数字位可装 / width one with sign leaves no digit position
ELSE
    nDigitsAvail := nWUse;                     // 无符号：全部位可装数字 / no sign, every position carries a digit
END_IF

(*------------------------------------------------------------------------------
 * 段 4｜负域逐位分解（本件核心防错：-**不取绝对值**）
 *      Negative-domain digit decomposition, the absolute value is never taken
 *      nValue = -2147483648 取绝对值即回绕，故负值直接进负域、正值取反进负域
 *      ABS(-2147483648) wraps, so negatives stay negative and positives are negated
 *-----------------------------------------------------------------------------*)
IF nValue < 0 THEN
    nWork := nValue;                            // 已属负域，原样使用 / already negative, used as is
ELSE
    nWork := -nValue;                           // 正数升到负域，最大 2147483647 → -2147483647 无溢出 / positive moved to the negative domain, no overflow
END_IF

sDigits := '';                                  // 数字段清空 / digit segment cleared
IF nWork = 0 THEN
    sDigits     := MID(DL_DIGITS, DL_POS_ONE, DL_POS_ONE); // 零值特例：单个字符 '0' / zero special case, a single character
    nDigitCount := 1;                           // 零视为一位 / zero counts as one digit
END_IF

WHILE (nWork <> 0) AND (nGuard <= DL_GUARD_MAX) DO
    nDigit   := -(nWork MOD DL_TEN);            // 负域取模得 0~-9，取反得 0~9 / negative remainder negated into 0~9
    sDigitCh := MID(DL_DIGITS, DL_POS_ONE, DINT_TO_INT(nDigit) + DL_POS_ONE); // 数字 → 字符，查表不靠字符码算术 / digit to character through the table
    sDigits  := CONCAT(sDigitCh, sDigits);      // 前插，保证高位在前 / prepended so the most significant digit leads
    nDigitCount := nDigitCount + DL_POS_ONE;    // 位数累计 / digit count incremented
    nWork    := nWork / DL_TEN;                 // 向零整除，负域同样正确 / truncating division, correct in the negative domain
    nGuard   := nGuard + DL_POS_ONE;            // 守卫累计，防死循环 / guard incremented, prevents a dead loop
END_WHILE

(*------------------------------------------------------------------------------
 * 段 5｜容量闸门（装不下就拒绝，绝不输出半截数字）
 *      Capacity gate: refuse when it does not fit, never emit a truncated number
 *-----------------------------------------------------------------------------*)
IF (nDigitCount > nDigitsAvail) OR (nDigitCount > DL_DIGIT_MAX) OR (nGuard > DL_GUARD_MAX) THEN
    eErr     := 16#0001_03A8;                   // 故障级：宽度不足，拒绝编码 / fault: insufficient width, encoding refused
    bError   := TRUE;                           // 置故障标志 / raise the fault flag
    bValid   := FALSE;                          // 结果不可用 / result unusable
    sField   := '';                             // 字段保持空串 / field stays empty
    uFieldLen := 0;                             // 写入长度保持 0 / written length stays zero
    FC_DL_IntToFixedField := FALSE;             // 返回失败 / return failure
    RETURN;                                     // 早退路径已统一后处理 / the early exit is fully post-processed
END_IF

(*------------------------------------------------------------------------------
 * 段 6｜填充段构造（个数 = 可用位 − 实际位数，恒非负）
 *      Pad segment build: available positions minus actual digits, never negative
 *-----------------------------------------------------------------------------*)
nPadCount := nDigitsAvail - nDigitCount;        // 段 5 已保证 nDigitCount ≤ nDigitsAvail / guaranteed non-negative by segment five
sPad      := '';                                // 填充段清空 / pad segment cleared
nGuard    := 0;                                 // 守卫复用前先清零 / guard cleared before reuse
WHILE (nPadCount > 0) AND (nGuard <= DL_W_MAX) DO
    IF bZeroPad THEN
        sPad := CONCAT(sPad, DL_PAD_ZERO);      // 零填充 / zero padding
    ELSE
        sPad := CONCAT(sPad, DL_PAD_SPACE);     // 空格填充 / space padding
    END_IF
    nPadCount := nPadCount - DL_POS_ONE;        // 剩余个数递减 / remaining count decremented
    nGuard    := nGuard + DL_POS_ONE;           // 守卫累计，上界为宽度上限 / guard bounded by the width limit
END_WHILE

(*------------------------------------------------------------------------------
 * 段 7｜符号段与拼装（对齐口径见头注释）
 *      Sign segment and assembly, alignment per the header rules
 *-----------------------------------------------------------------------------*)
IF bNeedSign THEN
    IF bNeg THEN
        sSign := DL_SIGN_MINUS;                 // 负号 / minus sign
    ELSE
        sSign := DL_SIGN_PLUS;                  // 强制正号 / forced plus sign
    END_IF
ELSE
    sSign := '';                                // 无符号段 / no sign segment
END_IF

IF bNeedSign AND bZeroPad THEN
    sField := CONCAT(sSign, CONCAT(sPad, sDigits)); // 零填充：符号贴最左 -0000042 / zero pad, sign on the far left
ELSE
    sField := CONCAT(sPad, CONCAT(sSign, sDigits)); // 空格填充：符号紧贴数字      -42 / space pad, sign next to the digits
END_IF

(*------------------------------------------------------------------------------
 * 段 8｜长度复检与出口（结构性不可能命中，纯防御纵深，R94 统一后处理）
 *      Length recheck and exit, structurally unreachable, pure defense in depth
 *-----------------------------------------------------------------------------*)
IF LEN(sField) <> nWUse THEN
    eErr     := 16#0001_03A8;                   // 复检不符：按同一故障码拒绝（不新增码位，R90） / recheck mismatch, same fault code, no new code
    bError   := TRUE;                           // 置故障标志 / raise the fault flag
    bValid   := FALSE;                          // 结果不可用 / result unusable
    sField   := '';                             // 字段回空，绝不交出不完整字段 / field emptied, never hand out an incomplete one
    uFieldLen := 0;                             // 写入长度回 0 / written length back to zero
    FC_DL_IntToFixedField := FALSE;             // 返回失败 / return failure
    RETURN;
END_IF

uFieldLen := INT_TO_UINT(nWUse);                // 写入字符数 = 生效宽度 / written length equals the effective width
bValid    := TRUE;                              // 结果可用 / result usable
FC_DL_IntToFixedField := TRUE;                  // 编码成功 / encoding succeeded
END_FUNCTION

(* ---- FC_DL_InvSqrtApprox.st ---- *)
// FC_DL_InvSqrtApprox v1.0.0
(*==============================================================================
 * 功能描述: 平方根倒数 1/sqrt(x) 快速近似。先按 4 倍缩放把自变量归一到 [1,4)，
 *           线性初值后牛顿迭代 4 次（残差 < 0.1%），再按缩放级数还原；缩放循环带
 *           128 步守护（R3 三族开闭词配对口径）；x <= 0 或非有限防御返回 0 并置
 *           bValid=FALSE。
 * 接口契约: 输入 fX，域 > 0 [无量纲]；输出 bValid 回执，返回 1/sqrt(x) 近似值。
 * 修订历史: 2026-11-23  v1.0.0  R74 首版
 *==============================================================================*)

FUNCTION FC_DL_InvSqrtApprox : REAL
VAR_INPUT
    fX : REAL := 1.0;   // 自变量，域 > 0 [无量纲] / Argument, domain > 0
END_VAR
VAR_OUTPUT
    bValid : BOOL;      // 结果有效回执 [-] / Result validity receipt
END_VAR
VAR CONSTANT
    DL_ISA_EPS : REAL := 1.0E-6;   // 判零容差 [无量纲] / Zero-test epsilon
END_VAR
VAR
    fScaled : REAL;     // 缩放后自变量（落在 [1,4)）[无量纲] / Scaled argument in [1,4)
    fY      : REAL;     // 牛顿迭代工作值 [无量纲] / Newton iteration working value
    nScale  : INT;      // 4 倍缩放级数 [级] / Scaling stages of factor four
    nGuard  : INT;      // 缩放循环守护计数 [步] / Scaling loop guard
END_VAR

(* —— 段 0：全路径赋值缺省（无效安全侧） —— *)
bValid := FALSE;                             // 有效回执预清 / Validity preset
FC_DL_InvSqrtApprox := 0.0;                  // 返回值缺省零 / Result default zero

(* —— 段 1：域闸与非有限闸 —— *)
IF fX <> fX THEN                             // NaN 自反判（判等禁令唯一例外） / NaN self-reflexive test
    RETURN;                                  // 无效返回零 / Invalid, return zero
END_IF
IF fX < DL_ISA_EPS THEN                      // 非正域拦截（含判零容差） / Non-positive domain intercepted
    RETURN;                                  // 无效返回零 / Invalid, return zero
END_IF
IF fX >= 3.0E38 THEN                         // 近 Inf 幅值闸 / Near-Inf magnitude gate
    RETURN;                                  // 无效返回零 / Invalid, return zero
END_IF

(* —— 段 2：4 倍缩放归一到 [1,4)（守护 128 步防死循环，R3 配对口径） —— *)
fScaled := fX;                               // 缩放工作值装载 / Scaled value seeded
nScale := 0;                                 // 缩放级数清零 / Stage count cleared
nGuard := 0;                                 // 守护计数清零 / Guard cleared
WHILE (fScaled >= 4.0) AND (nGuard < 128) DO // 大于等于 4 连续除 4 / Divide by four while at or above four
    fScaled := fScaled / 4.0;                // 除以 4（缩放一级） / Divide by four
    nScale := nScale + 1;                    // 级数递增 / Stage increments
    nGuard := nGuard + 1;                    // 守护递增 / Guard increments
END_WHILE                                    // WHILE 闭合（配对断言） / WHILE closed, pairing asserted

(* —— 段 3：线性初值 + 牛顿迭代 4 次（[1,4) 域内残差 < 0.1%） —— *)
fY := 0.95 - 0.15 * fScaled;                 // 线性初值（域内偏差 <= 30%） / Linear seed, deviation at most thirty percent
fY := fY * (3.0 - fScaled * fY * fY) / 2.0;  // 牛顿第 1 次：y*(3-x*y²)/2 / Newton iteration one
fY := fY * (3.0 - fScaled * fY * fY) / 2.0;  // 牛顿第 2 次 / Newton iteration two
fY := fY * (3.0 - fScaled * fY * fY) / 2.0;  // 牛顿第 3 次 / Newton iteration three
fY := fY * (3.0 - fScaled * fY * fY) / 2.0;  // 牛顿第 4 次 / Newton iteration four

(* —— 段 4：按缩放级数还原（每级乘 0.5，级数由守护上界钳定） —— *)
WHILE (nScale > 0) AND (nGuard < 256) DO     // 还原循环（守护二次覆盖） / Restore loop, second guard
    fY := fY * 0.5;                          // 每级乘 0.5（除以 2 的逆缩放） / Multiply by a half per stage
    nScale := nScale - 1;                    // 级数递减 / Stage decrements
    nGuard := nGuard + 1;                    // 守护递增 / Guard increments
END_WHILE                                    // WHILE 闭合（配对断言） / WHILE closed, pairing asserted
FC_DL_InvSqrtApprox := fY;                   // 返回近似值 / Return the approximation
bValid := TRUE;                              // 有效回执 / Validity receipt

END_FUNCTION

(* ---- FC_DL_Kalman2DSmoother.st ---- *)
(*
  ==================================================================
  组件名 Component  : FC_DL_Kalman2DSmoother
  分类   Category   : DL_MathData
  复杂度 Complexity  : cx5
  版本   Version    : 1.0.0
  功能   Purpose    : 2D 常速模型稳态卡尔曼平滑（纯函数形态，状态由外部持有）。
                      输入本拍测量 (zX, zY) 与上拍状态 (x, y, vx, vy)、采样周期 dt、
                      过程噪声 q、量测噪声 r，按标量序贯近似输出更新后状态与位置
                      估计。协方差用标量稳态近似：位置增益 alpha = q·dt / (q·dt + r)，
                      速度增益 beta = alpha² / (2 - alpha)（alpha-beta 滤波器即稳态
                      二态卡尔曼，公开结果）；速度修正经 beta/dt 施加。
  来源   Source     : ROADMAP R56 池（与 FB_DL_KalmanFilter1D 分工：1D 标量 vs 2D 常速）
  溯源   Origin     : IEC 61131-3 标准语义的道莅防御性实现；稳态卡尔曼与 alpha-beta
                      滤波等价性为公开控制理论结果，clean-room 自研实现，未复制任何
                      闭源代码行。
  平台   Platform   : 纯 IEC 61131-3（LREAL 运算，无私有库、无幂运算符）
  作者   Author     : 道莅代码库 · PLC 编程专家（R56）
  ------------------------------------------------------------------
  边界 Boundary     :
                      一 本件为纯函数，无跨扫描周期状态驻留，协方差不外显（标量稳态
                         近似内嵌于增益解析式，属主边界）；
                      二 失败语义（R191 显式声明）：r <= 0 / dt <= 0 / q < 0 / 任一输入
                         非有限时，出口原样返回上拍状态并置 bInvalid（冻结保持）；
                      三 dt 下界 1.0E-6 防速度修正除零（beta/dt）；
                      四 无全局变量、无外部变量声明、无物理地址寻址、无定时器（纯函数）。
  输出契约 Output contract:
                      xN / yN / vxN / vyN 仅在 bInvalid = FALSE 时为更新后状态；
                      本件为纯函数，无跨扫描周期状态驻留。
  修订记录 Revision  :
    2026-11-20  v1.0.0  R56 首版（批 2 · 序号 6）
  ==================================================================
*)

FUNCTION FC_DL_Kalman2DSmoother : BOOL
VAR_INPUT
    zX : LREAL; // X 轴测量值 [长度单位] / X axis measurement [length unit]
    zY : LREAL; // Y 轴测量值 [长度单位] / Y axis measurement [length unit]
    x  : LREAL; // 上拍 X 位置估计 [长度单位] / previous X position estimate [length unit]
    y  : LREAL; // 上拍 Y 位置估计 [长度单位] / previous Y position estimate [length unit]
    vx : LREAL; // 上拍 X 速度估计 [长度每秒] / previous X velocity estimate [length per second]
    vy : LREAL; // 上拍 Y 速度估计 [长度每秒] / previous Y velocity estimate [length per second]
    dt : LREAL; // 采样周期 [秒]，域 大于零 / sample period [second], domain above zero
    q  : LREAL; // 过程噪声强度（每秒）[平方长度每秒] / process noise intensity per second [square length per second]
    r  : LREAL; // 量测噪声方差 [平方长度] / measurement noise variance [square length]
END_VAR
VAR_OUTPUT
    xN      : LREAL; // 更新后 X 位置估计 [长度单位] / updated X position estimate [length unit]
    yN      : LREAL; // 更新后 Y 位置估计 [长度单位] / updated Y position estimate [length unit]
    vxN     : LREAL; // 更新后 X 速度估计 [长度每秒] / updated X velocity estimate [length per second]
    vyN     : LREAL; // 更新后 Y 速度估计 [长度每秒] / updated Y velocity estimate [length per second]
    bInvalid: BOOL;  // 输入无效，出口原样返回上拍状态 [-] / the input is void, the outlet returns the previous state unchanged
END_VAR
VAR
    _bFin  : BOOL := FALSE;  // 九个输入全部有限 [-] / all nine inputs are finite
    _fDt   : LREAL := 0.0;   // 钳定后的采样周期 [秒] / the clamped sample period [second]
    _fQdt  : LREAL := 0.0;   // 过程噪声强度乘周期 [平方长度] / process noise times the period
    _fAlp  : LREAL := 0.0;   // 位置增益 alpha [无量纲] / the position gain alpha
    _fBta  : LREAL := 0.0;   // 速度增益 beta [无量纲] / the velocity gain beta
    _fPx   : LREAL := 0.0;   // X 轴位置预测 [长度单位] / the X position prediction
    _fPy   : LREAL := 0.0;   // Y 轴位置预测 [长度单位] / the Y position prediction
    _fIx   : LREAL := 0.0;   // X 轴新息 [长度单位] / the X innovation
    _fIy   : LREAL := 0.0;   // Y 轴新息 [长度单位] / the Y innovation
END_VAR

// 段 1｜非有限闸（R151 全覆盖）与参数域闸 / segment 1, finiteness gate over every input and the parameter domain gate
_bFin := (zX = zX) AND ((zX - zX) = (zX - zX)) AND (zY = zY) AND ((zY - zY) = (zY - zY)) AND (x = x) AND ((x - x) = (x - x)) AND (y = y) AND ((y - y) = (y - y)) AND (vx = vx) AND ((vx - vx) = (vx - vx)) AND (vy = vy) AND ((vy - vy) = (vy - vy)) AND (dt = dt) AND ((dt - dt) = (dt - dt)) AND (q = q) AND ((q - q) = (q - q)) AND (r = r) AND ((r - r) = (r - r)); // 九输入有限性 / finiteness of all nine inputs
IF (NOT _bFin) OR (dt <= 0.0) OR (r <= 0.0) OR (q < 0.0) THEN // 输入无效或参数越域 / the input is void or a parameter is out of domain
    xN := x;   // 冻结保持：原样返回上拍状态（R191 显式声明）/ frozen hold, the previous state passes through unchanged
    yN := y;   // 冻结保持 / frozen hold
    vxN := vx; // 冻结保持 / frozen hold
    vyN := vy; // 冻结保持 / frozen hold
    bInvalid := TRUE; // 置无效标志 / raise the invalid flag
    FC_DL_Kalman2DSmoother := FALSE; // 函数返回失败 / the function returns failure
    RETURN; // 早退 / early return
END_IF

// 段 2｜稳态增益计算（标量近似） / segment 2, the steady state gains by the scalar approximation
_fDt := dt; // 周期直通 / the period passes through
IF _fDt < 1.0E-6 THEN // 周期过小 / the period is too small
    _fDt := 1.0E-6; // 抬到下限，防速度修正除零 / raised against the velocity divisor
END_IF
_fQdt := q * _fDt; // 过程噪声强度乘周期 / the process noise times the period
_fAlp := _fQdt / (_fQdt + r); // 位置增益，除子为 q·dt + r 已证 > 0 / the position gain, the divisor is proven positive
_fBta := _fAlp * _fAlp / (2.0 - _fAlp); // 速度增益，除子 2 - alpha 已证 > 1（alpha < 1 结构性成立）/ the velocity gain, the divisor is proven above one since alpha is structurally below one

// 段 3｜X 轴预测与更新 / segment 3, the X axis prediction and update
_fPx := x + vx * _fDt; // 常速位置预测 / the constant velocity position prediction
_fIx := zX - _fPx; // 新息 / the innovation
xN := _fPx + _fAlp * _fIx; // 位置更新 / the position update
vxN := vx + (_fBta / _fDt) * _fIx; // 速度更新（除子已钳下限）/ the velocity update with the proven divisor

// 段 4｜Y 轴预测与更新 / segment 4, the Y axis prediction and update
_fPy := y + vy * _fDt; // 常速位置预测 / the constant velocity position prediction
_fIy := zY - _fPy; // 新息 / the innovation
yN := _fPy + _fAlp * _fIy; // 位置更新 / the position update
vyN := vy + (_fBta / _fDt) * _fIy; // 速度更新（除子已钳下限）/ the velocity update with the proven divisor

bInvalid := FALSE; // 有效标志 / the valid flag
FC_DL_Kalman2DSmoother := TRUE; // 函数返回成功 / the function returns success
END_FUNCTION

(* ---- FC_DL_LagrangeInterp.st ---- *)
(*==============================================================================
 * 组件名称 (Component)  : FC_DL_LagrangeInterp
 * 所属子库 (Sublibrary) : DL_MathData
 * 当前版本 (Version)    : 1.0.0
 * 兼容性   (Platform)   : CODESYS 3.5+ / TwinCAT 3 / 汇川 InoProShop / 施耐德 Machine Expert
 *                         仅依赖 Standard.library（LOWER_BOUND / UPPER_BOUND / ABS），零厂商私有库
 * 功能描述 (Function)   : 小样本拉格朗日插值原语：对 2 ≤ n ≤ 8 个散点 (aX[i], aY[i])，
 *                         以拉格朗日基函数求单点插值
 *                           fYq = Σ_i aY[i] × Π_{j≠i} (fXq - aX[j]) / (aX[i] - aX[j])
 *                         适用 2~8 点传感器标定曲线（如 NTC 温度、压力标定）的非线性插值。
 * 接口     (Interface)  : 输入 aX 横坐标数组（变长数组，按引传）、aY 纵坐标数组（变长数组，
 *                         按引传）、fXq 查询横坐标；引用输出 bValid 有效标志
 *                         （REFERENCE TO BOOL，当拍写回）；返回值 = 插值结果
 *                         （bValid=FALSE 时返回 0）。
 * 边界     (Boundary)   : ① **属主边界（写死）：本件只做一次静态散点求值，不装载标定表、
 *                         不缓存系数、不做外推告警**；标定表管理由调用方负责。
 *                         ② 拒算条件（任一成立返回 0 且 bValid=FALSE）：点数 < 2、两数组
 *                         长度不一致、fXq 非有限、任一点非有限（NaN 自不等 x<>x、Inf 用
 *                         (x-x)<>0 口径）、查重节点（ABS(aX[i]-aX[j]) < 节点容差，分母趋零，
 *                         浮点禁 = 判等，R28）。
 *                         ③ 点数超上限（8）按**截断语义**处理：只取前 8 点求值并在
 *                         bValid=TRUE 下照常返回，截断行为写死于此，调用方按需自校点数。
 *                         ④ 节点容差提为 VAR CONSTANT（禁魔法数）；无样条连续性要求的小
 *                         样本域适用，需要 C2 连续时改用 `FC_DL_CubicSplineInterp`。
 *                         ⑤ 变长数组仅入 VAR_IN_OUT（ARRAY[*] 传参域限定），实际上下界由
 *                         LOWER_BOUND/UPPER_BOUND 取得，不假设 0 起始。
 *                         ⑥ 零全局耦合（无 GVL / 无 VAR_EXTERNAL / 无物理地址）。
 * 分工声明 (Scope)      : 与 `FC_DL_CubicSplineInterp` 分工：无样条连续性要求的小样本多项式
 *                         插值（本件）≠ 三次样条 C2 连续插值（那件），实现独立不复制；
 *                         与 `FC_DL_MultiPointLinear` 分工：多项式过点 ≠ 分段线性。
 * 来源标签 (Source Tag) : T2-1 LGF · Math 数学子族（公开数学定义 clean-room，拉格朗日
 *                         基函数为教科书公开公式，零代码行复制）
 * 码表     (Codes)      : 本件不占用任何全局数字码位。出口为 LREAL 插值 + BOOL 有效标志；
 *                         数字码位待主控收口阶段统一派号。
 * 红线自检 (Redline)    : R1 ✓ 零 GVL/VAR_EXTERNAL ｜ R2 ✓ 零 %I/%Q/%M ｜ R3 ✓ 纯 IEC 61131-3
 *                         R4 ✓ 节点容差查重 + 非有限前置剔除 + 点数上限钳位 ｜ R5 ✓ 声明逐行同行双语注释
 *                         R6 N/A（纯函数无状态机） ｜ R7 N/A（无实例调用）
 * 修订历史 (Revision)   : 2026-11-20  v1.0.0  R48 首版（批次 1 · 序号 3）
 *                         验收向量：2 点线性退化为直线；3 点过三抛物线；重节点拒算；
 *                         9 点输入按前 8 点截断求值。
 *==============================================================================*)

FUNCTION FC_DL_LagrangeInterp : LREAL
VAR_IN_OUT
    aX : ARRAY[*] OF LREAL;    // 节点横坐标数组（散点，须互异），单位随横轴 [横轴单位] / Node abscissae, distinct
    aY : ARRAY[*] OF LREAL;    // 节点纵坐标数组，单位随纵轴 [纵轴单位] / Node ordinates
END_VAR
VAR_INPUT
    fXq    : LREAL;                 // 查询横坐标（允许落在节点域外，外推不告警） [横轴单位] / Query abscissa, extrapolation allowed
    bValid : REFERENCE TO BOOL;     // 有效标志（引用传参；FALSE=拒算） [-] / Validity flag, by-reference, FALSE when rejected
END_VAR
VAR
    nLo    : DINT;                  // aX 数组实际下界索引 / Lower index of aX
    nHiX   : DINT;                  // aX 数组实际上界索引 / Upper index of aX
    nHiY   : DINT;                  // aY 数组实际上界索引 / Upper index of aY
    nCount : DINT;                  // 有效点数（截断后）/ Effective point count after truncation
    i      : DINT;                  // 基函数外层循环索引 / Outer basis loop index
    j      : DINT;                  // 基函数内层循环索引 / Inner basis loop index
    fYq    : LREAL;                 // 插值累加中间量 [纵轴单位] / Interpolation accumulator
    fTerm  : LREAL;                 // 单项基函数乘积中间量 [纵轴单位] / Single basis product term
END_VAR
VAR CONSTANT
    DL_LI_NMAX : DINT  := 8;        // 点数上限（2~8 小样本域） [点] / Point-count ceiling
    DL_LI_TOL  : LREAL := 1.0E-9;   // 查重节点容差（分母趋零闸） [横轴单位] / Duplicate-node tolerance
    DL_LI_EPS  : LREAL := 0.0;      // 非有限差值判零基准 [横轴单位] / Non-finite difference zero base
END_VAR

bValid := FALSE;                                       // 缺省拒算 / Default: invalid
FC_DL_LagrangeInterp := 0.0;                           // 拒算返回 0 / Rejected returns zero
nLo    := LOWER_BOUND(aX, 1);                          // aX 实际下界 / Actual lower bound of aX
nHiX   := UPPER_BOUND(aX, 1);                          // aX 实际上界 / Actual upper bound of aX
nHiY   := UPPER_BOUND(aY, 1);                          // aY 实际上界 / Actual upper bound of aY
IF (nHiX - nLo) <> (nHiY - LOWER_BOUND(aY, 1)) THEN
    RETURN;                                            // 两数组长度不一致：拒算 / Length mismatch: reject
END_IF
nCount := nHiX - nLo + 1;                              // 原始点数 / Raw point count
IF (fXq <> fXq) OR ((fXq - fXq) <> DL_LI_EPS) THEN
    RETURN;                                            // 查询值非有限（NaN/Inf）：拒算 / Non-finite query: reject
END_IF
IF nCount < 2 THEN
    RETURN;                                            // 点数不足 2：拒算 / Fewer than two points: reject
END_IF
IF nCount > DL_LI_NMAX THEN
    nCount := DL_LI_NMAX;                              // 超上限截断语义：只取前 8 点（声明于头注释③） / Truncate to ceiling per header clause 3
END_IF
nHiX := nLo + nCount - 1;                              // 截断后有效上界 / Effective upper bound after truncation

FOR i := nLo TO nHiX DO
    IF (aX[i] <> aX[i]) OR ((aX[i] - aX[i]) <> DL_LI_EPS)
       OR (aY[i] <> aY[i]) OR ((aY[i] - aY[i]) <> DL_LI_EPS) THEN
        RETURN;                                        // 任一点非有限：整体拒算（R245）/ Any non-finite point: reject wholly
    END_IF
END_FOR
FOR i := nLo TO (nHiX - 1) DO
    FOR j := (i + 1) TO nHiX DO
        IF ABS(aX[i] - aX[j]) < DL_LI_TOL THEN
            RETURN;                                    // 查重节点命中（分母趋零）：拒算（R28 浮点禁 =）/ Duplicate nodes: reject
        END_IF
    END_FOR
END_FOR

fYq := 0.0;                                            // 插值累加器清零 / Clear accumulator
FOR i := nLo TO nHiX DO
    fTerm := aY[i];                                    // 单项从纵坐标出发 / Term starts from ordinate
    FOR j := nLo TO nHiX DO
        IF j <> i THEN
            fTerm := fTerm * (fXq - aX[j]) / (aX[i] - aX[j]);   // 基函数因子（分母已过查重闸）/ Basis factor, denominator gate-passed
        END_IF
    END_FOR
    fYq := fYq + fTerm;                                // 累加单项 / Accumulate term
END_FOR

FC_DL_LagrangeInterp := fYq;                           // 返回插值结果 / Return interpolated value
bValid := TRUE;                                        // 求值有效 / Result valid

END_FUNCTION

(* ---- FC_DL_LerpClamped.st ---- *)
(*
    FC_DL_LerpClamped —— 线性插值（t 域钳位，端点外不外推）
    ------------------------------------------------------------------
    组件名称  : FC_DL_LerpClamped
    分类      : DL_MathData / Interpolation
    前缀      : FC_DL_
    版本      : 1.0.0
    溯源      : 借鉴点 —— 数值分析中带参数域钳位的两点线性插值（lerp）语义，
                即 clamp 后的凸组合形式 y = a + (b - a) * clamp(t, 0, 1)；
                该形式在 t 超出 [0,1] 时**退回端点值**而不外推，是设定值过渡、
                配方插值、执行器软过渡的通行做法。
                clean-room 声明 —— 零代码行复制，只使用标准算术运算符与标准
                标准库函数 ABS；域闸 / 饱和 / 码位 / 双语文档全部自有。
                许可证 —— 本件 MIT；来源标签 self-std（道莅自有内规族），
                参考语义为公开数值方法常识，无第三方源码继承。
    平台      : 纯 IEC 61131-3，CODESYS 3.5 / TwinCAT 3 / InoProShop / Machine Expert 通用
    作者      : 道莅代码库 · PLC编程专家（R70 构建轮 · 批 1 · N2）
    ------------------------------------------------------------------
    功能说明  : 对端点 fA、fB 依参数 fT 做线性插值，fT 先钳到 [0,1]。
                「不外推」是本件与裸 lerp 的唯一语义差别：fT < 0 返回 fA，
                fT > 1 返回 fB，中间按凸组合。
                非有限闸（R272 逐项点名，含换算与限值）：fA / fB / fT 三入参
                全部纳入 NaN 自反判 + Inf 差值自反判 + 幅值 1E30 上界筛查；
                闸不通过时**结构早退**并返回安全缺省值 fA（端点 A 为稳态值，
                不是中间插值，避免故障时输出一个凭空构造的中间量）。
                凸组合实现口径（关键设计）：先算 fT 钳位值 fTc，再算
                差值 fB - fA，最后 fA + 差值 * fTc。差值可能超 LREAL 域，
                故对中间量做**结果非有限复检**：若委托乘法后结果非有限，
                按端点就近原则饱和到 fB 或 fA 并报信息级，绝不把 Inf 送下游。
                本件无除法（凸组合形式不带除法），故不存在除零面。
    错误码    : 16#0002_0111 入参非有限（NaN / Inf / 超幅值），返回 fA —— 故障级
                16#0002_0112 插值结果非有限，已饱和至端点 —— 信息级，值可用
    码位总账  : 16#0002_0111 用 ｜ 16#0002_0112 用
    状态机    : R6 N/A —— 纯函数无状态，无 CASE 可写，非法状态不可能出现
    边界与披露: 一 无定时器 / 无边沿实例 / 无数组下标，周期安全规则 N/A；
                二 零全局变量、零 VAR_EXTERNAL、零物理地址；
                三 bClamped 表示 fT 曾被钳位（含恰为 0 / 1 的边界情形，
                   判据为钳位前后是否同值，不含容差 —— 布尔判据非浮点判据，
                   但比较用差值容差口径以避开浮点直比）；
                四 结果非有限分支置「端点 + 信息级」而非故障级：饱和是防御
                   动作、值仍可用于下游限幅链路，R45 口径要求信息级不置 bError。
    修订记录  : 2026-11-22 v1.0.0 首次入库（R70 构建轮 · 批 1 · N2）
*)
FUNCTION FC_DL_LerpClamped : LREAL
VAR_INPUT
    fA : LREAL;                            (* 端点 A 的值，[工程单位] / the value at endpoint A *)
    fB : LREAL;                            (* 端点 B 的值，[工程单位] / the value at endpoint B *)
    fT : LREAL;                            (* 插值参数，[0..1] 为有效域，域外钳位 / the interpolation parameter, clamped to 0..1 *)
END_VAR
VAR_OUTPUT
    eErr     : UDINT;                      (* 错误码，0 = 正常 / the error id, 0 = ok *)
    bError   : BOOL;                       (* 故障标志，故障级码时 TRUE / the error flag, TRUE on fault level *)
    bValid   : BOOL;                       (* 返回值可用，故障级为 FALSE / the return usable, FALSE on fault level *)
    bClamped : BOOL;                       (* fT 曾被钳到 [0,1] 域内，[标志] / the parameter was clamped into 0..1 *)
    fTUsed   : LREAL;                      (* 实际参与运算的钳位后参数，[无量纲] / the clamped parameter actually used *)
END_VAR
VAR CONSTANT
    DL_LRP_FMAX : LREAL := 1.0E30;         (* 非有限筛查幅值上限，[工程单位] / the finiteness screening cap *)
    DL_LRP_TOL  : LREAL := 1.0E-12;        (* 参数域钳位的比较容差，[无量纲] / the clamp comparison tolerance *)
END_VAR
VAR
    _fT  : LREAL;                          (* 钳位后的参数（内部中间量），[无量纲] / the clamped parameter, an internal temporary *)
    _fD  : LREAL;                          (* 端点差值 fB - fA（内部中间量），[工程单位] / the endpoint delta, an internal temporary *)
    _fY  : LREAL;                          (* 插值结果（内部中间量），[工程单位] / the interpolation result, an internal temporary *)
END_VAR

// 段 1｜返回值与状态预置（四段式第一段）/ segment 1, preset the return and the status
FC_DL_LerpClamped := fA;               // 故障缺省返回端点 A（稳态值）/ the fault default is endpoint A, a steady value
eErr     := 0;                         // 预置无错误 / preset no error
bError   := FALSE;                     // 预置无故障 / preset no fault
bValid   := FALSE;                     // 预置不可用，过闸后置位 / preset unusable, set TRUE after the gates
bClamped := FALSE;                     // 预置未钳位 / preset not clamped
fTUsed   := 0.0;                       // 预置参数出口零值 / preset the parameter outlet to zero

// 段 2｜三入参非有限闸（NaN 自反判 + Inf 差值自反判 + 幅值上界，R272 逐项点名）/ segment 2, the finiteness gate
IF (fA <> fA) OR ((fA - fA) <> 0.0) OR (ABS(fA) > DL_LRP_FMAX) THEN   // 端点 A 非有限 / endpoint A non finite
    eErr   := 16#0002_0111;            // 故障级：入参非有限 / fault level: a non finite input
    bError := TRUE;                    // R45 配对置故障标志 / paired with the code
    bValid := FALSE;                   // 返回值不可用 / the return is unusable
    RETURN;                            // 结构早退 / structural exit
END_IF
IF (fB <> fB) OR ((fB - fB) <> 0.0) OR (ABS(fB) > DL_LRP_FMAX) THEN   // 端点 B 非有限 / endpoint B non finite
    eErr   := 16#0002_0111;            // 故障级：入参非有限 / fault level: a non finite input
    bError := TRUE;                    // R45 配对 / paired with the code
    bValid := FALSE;                   // 返回值不可用 / the return is unusable
    RETURN;                            // 结构早退 / structural exit
END_IF
IF (fT <> fT) OR ((fT - fT) <> 0.0) OR (ABS(fT) > DL_LRP_FMAX) THEN   // 插值参数非有限 / the parameter non finite
    eErr   := 16#0002_0111;            // 故障级：入参非有限 / fault level: a non finite input
    bError := TRUE;                    // R45 配对 / paired with the code
    bValid := FALSE;                   // 返回值不可用 / the return is unusable
    RETURN;                            // 结构早退 / structural exit
END_IF

// 段 3｜参数域闸：t 钳到 [0,1]，域外不外推 / segment 3, the parameter domain clamp
_fT := fT;                             // 取参数原值 / take the raw parameter
IF fT < 0.0 THEN                       // 低于下域界 / under the lower domain edge
    _fT := 0.0;                        // 钳到 0，输出退回端点 A / clamp to zero, fall back to endpoint A
    bClamped := TRUE;                  // 记录已钳位 / record the clamp
ELSIF fT > 1.0 THEN                    // 高于上域界 / over the upper domain edge
    _fT := 1.0;                        // 钳到 1，输出退回端点 B / clamp to one, fall back to endpoint B
    bClamped := TRUE;                  // 记录已钳位 / record the clamp
END_IF
fTUsed := _fT;                         // 参数出口（钳位后真值）/ the parameter outlet, the clamped value

// 段 4｜凸组合委托：端点 + 差值 × 钳位参数（无除法，无除零面）/ segment 4, the convex combination kernel
_fD := fB - fA;                        // 端点差值，[工程单位] / the endpoint delta
_fY := fA + _fD * _fT;                 // 插值结果（委托 `+` 与 `*`）/ the interpolation result, delegated
IF (_fY <> _fY) OR ((_fY - _fY) <> 0.0) THEN   // 结果非有限（差值超域所致）/ the result came out non finite
    IF (ABS(_fT - 1.0) <= DL_LRP_TOL) THEN     // 参数贴 1 侧 / the parameter sits at the upper edge
        FC_DL_LerpClamped := fB;       // 饱和到端点 B / saturate to endpoint B
    ELSE                               // 参数在域内或贴 0 侧 / the parameter inside or at the lower edge
        FC_DL_LerpClamped := fA;       // 饱和到端点 A / saturate to endpoint A
    END_IF
    eErr   := 16#0002_0112;            // 信息级：结果非有限已饱和 / info level: the result was saturated
    bError := FALSE;                   // 信息级不置故障（R45）/ info level never raises the fault flag
    bValid := TRUE;                    // 端点值可用 / the endpoint value is usable
    RETURN;                            // 出口 / exit
END_IF

// 段 5｜域内正常出口 / segment 5, the in-domain outlet
FC_DL_LerpClamped := _fY;              // 域内插值结果 / the in-domain interpolation result
bError := FALSE;                       // 本路径无故障 / no fault on this path
bValid := TRUE;                        // 结果可用 / the result is usable
END_FUNCTION

(* ---- FC_DL_LimitEx.st ---- *)
(*
    FC_DL_LimitEx —— 三输入限幅泛型防御包装（REAL 域）
    ------------------------------------------------------------------
    分类      : DL_MathData / MinMax
    前缀      : FC_DL_
    版本      : 1.0.0
    溯源      : IEC 61131-3 标准语义的道莅防御性实现
                （内部委托平台内建函数，外围统一错误码/钳位/双语文档；
                  未复制任何闭源厂商源码，参考实现仅限 MIT/Apache 许可）
    平台      : 纯 IEC 61131-3，CODESYS / TwinCAT / InoProShop 通用
    作者      : 道莅代码库 · PLC编程专家（R16）
    ------------------------------------------------------------------
    功能说明  : 三输入限幅：将 fIn 限制在 [fMin, fMax] 区间内，比较与选择
                运算用 IF/ELSE 实现（IEC LIMIT 语义），不重实现任何数学内核；
                防御性交换声明：fMin > fMax 时自动交换上下限并置信息级 16#0001_01DE
                （bError=FALSE、bValid=TRUE，保证限幅区间恒有效）；
                三输入任一非有限（NaN 或 ±INF）判为故障级 16#0001_02BB，
                返回 0.0 且 bValid=FALSE（非有限值参与限幅语义未定义，一律拦截）；
                钳位方向：域内值钳至 [下限, 上限] 区间（LIMIT 本义钳位）；
                ±INF 采用平台安全幅值比较判定（阈值高于 REAL 最大有限值 3.402823E38），NaN 用自不等判定。
    错误码    : 16#0001_02BB 任一输入非有限（NaN 或 ±INF）——故障级，返回 0.0
                16#0001_01DE 上下限倒置，已自动交换（fMin 与 fMax 互换）——信息级，正常防御
                16#0001_01DF 预留禁用（信息级，不得挪用）
                16#0001_02BC 预留禁用（故障级，不得挪用）
                16#0001_02BD 预留禁用（故障级，不得挪用）
    状态机    : R6 标注 N/A —— 本组件为纯函数无顺序状态机，无 CASE 可写，非法状态不可能出现，故以本节说明替代 ELSE 兜底
    修订记录  : 2026-11-16 v1.0.0 首次入库（R16）
*)
FUNCTION FC_DL_LimitEx : REAL
VAR_INPUT
    fMin : REAL; // 限幅下限 [无量纲]，大于上限时自动交换 / lower limit, auto-swapped when greater than upper
    fIn  : REAL; // 限幅输入值 [无量纲] / value to be limited
    fMax : REAL; // 限幅上限 [无量纲]，小于下限时自动交换 / upper limit, auto-swapped when less than lower
END_VAR
VAR_OUTPUT
    eErr   : UDINT; // 错误码，0=正常 / error id, 0=ok
    bError : BOOL;  // 是否出错，eErr 非 0 时为 TRUE / error flag, TRUE when eErr is nonzero
    bValid : BOOL;  // 输出是否有效可用 / output valid flag
END_VAR
VAR CONSTANT
    DL_REAL_INF_GUARD : LREAL := 4.0E38; // REAL 域 ±INF 判定阈值，高于 REAL 最大有限值 3.402823E38 [无量纲] / REAL +/-INF guard above max finite REAL 3.402823E38
END_VAR
VAR
    fLo    : REAL; // 整备后的限幅下限 [无量纲] / prepared lower bound
    fHi    : REAL; // 整备后的限幅上限 [无量纲] / prepared upper bound
    bBad   : BOOL; // 任一输入非有限判定结果 / non-finite detection result of any input
END_VAR

// 段 1｜返回值与错误状态预置 / segment 1, preset return value and error status
FC_DL_LimitEx := 0.0; // 故障缺省返回 0 [无量纲] / fault default returns 0
eErr   := 0;     // 预置无错误 / preset no error
bError := FALSE; // 预置无故障 / preset no fault
bValid := FALSE; // 预置无效，通过防御闸后置位 / preset invalid, set TRUE after guard passes

// 段 2｜三输入非有限防御闸 / segment 2, three-input non-finite guard
bBad := (fMin <> fMin) OR (fMin > DL_REAL_INF_GUARD) OR (fMin < -DL_REAL_INF_GUARD)
     OR (fIn  <> fIn)  OR (fIn  > DL_REAL_INF_GUARD) OR (fIn  < -DL_REAL_INF_GUARD)
     OR (fMax <> fMax) OR (fMax > DL_REAL_INF_GUARD) OR (fMax < -DL_REAL_INF_GUARD); // 三输入非有限判定（NaN 自不等 + 安全幅值判 ±INF） [无量纲] / all three inputs non-finite check (NaN by self-inequality, +/-INF by safe magnitude)
IF bBad THEN
    FC_DL_LimitEx := 0.0;     // 故障级返回 0 [无量纲] / fault level returns 0
    eErr   := 16#0001_02BB;   // 非有限输入故障码 / non-finite input fault id
    bError := TRUE;           // 置故障标志 / set fault flag
    bValid := FALSE;          // 输出无效 / output invalid
    RETURN;                   // 立即返回 / immediate return
END_IF

// 段 3｜上下限整备（含防御性交换） / segment 3, bound preparation with defensive swap
IF fMin > fMax THEN
    fLo := fMax; // 倒置时下限取原上限 / swapped: lower takes original upper
    fHi := fMin; // 倒置时上限取原下限 / swapped: upper takes original lower
    eErr := 16#0001_01DE; // 信息级：上下限倒置已自动交换 / info level: bounds inverted, auto-swapped
ELSE
    fLo := fMin; // 正常序下限直通 / normal order, lower passes through
    fHi := fMax; // 正常序上限直通 / normal order, upper passes through
END_IF

// 段 4｜主体限幅计算（末段） / segment 4, main limiting calculation (final)
IF fIn < fLo THEN
    FC_DL_LimitEx := fLo; // 低于下限，钳至下限 / below lower bound, clamp to lower
ELSIF fIn > fHi THEN
    FC_DL_LimitEx := fHi; // 高于上限，钳至上限 / above upper bound, clamp to upper
ELSE
    FC_DL_LimitEx := fIn; // 区间内直通 / inside bounds, pass through
END_IF
bError := FALSE; // 信息级交换不置故障，故障分支已提前返回 / info-level swap never raises fault, fault branch has returned
bValid := TRUE;  // 域内或限幅输出均有效可用 / in-domain or limited output is valid
END_FUNCTION

(* ---- FC_DL_LinearRegression2Var.st ---- *)
(*
  FC_DL_LinearRegression2Var  —  二元最小二乘回归（3x3 正规方程）/ Two-variable least-squares linear regression
  分类 Category : DL_MathData
  码位 Code     : 16#05_0_02
  版本 Version  : 1.0.0
  来源 Source   : t2-1-lgf-math — IEC 61131-3 标准语义的道莅防御性实现
  溯源 Origin   : clean-room 实现，最小二乘正规方程公开数学语义，未复制任何源码行（命名对齐既有件 FC_DL_LinearScale）
  功能 Function : 1) 由 (x1, x2, y) 样本集解 3x3 正规方程（Cramer 法则），输出双斜率 fK1/fK2、截距 fB 与拟合优度 fR2；
                  2) 共线性判据：|r12| 越限即判「不可辨识」，不输出斜率（防病态解误导）；
                  3) 每个样本做非有限值（NaN/Inf）预筛，任一非法则整批无效。
  边界 Boundary : ① nSampleCount < 4 判样本不足置码（3 参数 3 方程不可给 R²），不进入求解；
                  ② nSampleCount 超数组上界判组态错置码（防越界，循环带上限守卫）；
                  ③ |r12| > fCollinearLimit 置 bIdentifiable := FALSE 且斜率/截距/R² 全 0（不给看似可信数字）；
                  ④ 行列式 |det| < 1E-12 判退化置 bDegenerate；
                  ⑤ SStot 近零（y 全等）时 R² 置 0 并置信息码（防除零）；
                  ⑥ 解除式自证：bIdentifiable/bDegenerate 为每调用重算量，下一调用条件消失即自动解除（无锁存）。
  依赖 Depends  : 仅 Standard.library（ABS/SQRT）；参考对齐 FC_DL_LinearScale（已注册，仅命名体例）
  码表 Error codes（本件格 05_0_02，子码步进 +0x100）:
    16#0005_0102 信息级：共线性越限，判不可辨识（bIdentifiable = FALSE）
    16#0005_0202 故障级：样本不足 nSampleCount < 4 或超数组上界
    16#0005_0302 故障级：样本含非有限值（NaN/Inf），整批无效
    16#0005_0402 故障级：正规方程退化（行列式 |det| < 1E-12）
    16#0005_0502 信息级：SStot 近零，R² 置 0（y 全等，拟合优度无定义）

  修订历史 Revision :
    2026-11-18  v1.0.0  R38 首版
*)

FUNCTION FC_DL_LinearRegression2Var : BOOL
VAR_INPUT
    afX1           : ARRAY[0..63] OF REAL;   // 样本 x1 组 [工程量] / Sample array x1
    afX2           : ARRAY[0..63] OF REAL;   // 样本 x2 组 [工程量] / Sample array x2
    afY            : ARRAY[0..63] OF REAL;   // 样本 y 组 [工程量] / Sample array y
    nSampleCount   : INT;                    // 有效样本数 [个]，域 4..64 / Valid sample count
    fCollinearLimit: REAL := 0.995;          // 共线性判据上限 |r12|，域 0..1 / Collinearity limit on |r12|
END_VAR
VAR_OUTPUT
    fK1            : REAL;                   // 回归斜率 1 [y 单位/x1 单位] / Regression slope k1
    fK2            : REAL;                   // 回归斜率 2 [y 单位/x2 单位] / Regression slope k2
    fB             : REAL;                   // 回归截距 [y 单位] / Regression intercept
    fR2            : REAL;                   // 拟合优度 R² [无量纲，0..1] / Coefficient of determination
    bIdentifiable  : BOOL;                   // 可辨识标志（共线性未越限）/ Identifiable flag
    bDegenerate    : BOOL;                   // 正规方程退化标志 / Degenerate normal-equation flag
    nErrId         : UDINT;                  // 事件码，0 = 无事件 / Event code, 0 = none
END_VAR
VAR
    rN, rSx1, rSx2, rSy      : LREAL;        // 计数与一次矩累加器 / Count and first-moment accumulators
    rS11, rS22, rS12         : LREAL;        // 二次矩累加器 / Second-moment accumulators
    rS1y, rS2y, rSyy         : LREAL;        // 交叉矩累加器 / Cross-moment accumulators
    rM1, rM2, rMy            : LREAL;        // 均值 x1/x2/y / Means of x1, x2 and y
    rV1, rV2, rC12           : LREAL;        // 方差与协方差（中心化）/ Central variances and covariance
    rR12, rDet, rDen         : LREAL;        // 相关系数/行列式/求根分母 / Correlation, determinant, solve denominator
    rSsTot, rSsRes, rYhat    : LREAL;        // 总平方和/残差平方和/拟合值 / Total SS, residual SS, fitted value
    rDx1, rDx2, rDy          : LREAL;        // 单样本临时量（LREAL 宽域防累加误差）/ Per-sample scratch
    bFin                     : BOOL;         // 非有限值筛查标志 / Non-finite screening flag
    k                        : INT;          // 循环计数器 / Loop counter
END_VAR
VAR CONSTANT
    nMaxSmp   : INT    := 64;      // 数组上界 [个] / Array upper bound
    rDetFloor : LREAL  := 1.0E-12; // 行列式退化阈值 / Degenerate determinant threshold
    rSsFloor  : LREAL  := 1.0E-12; // SStot 近零阈值 / Near-zero SStot threshold
    rFinLim   : LREAL  := 1.0E30;  // 非有限值筛查幅值上限 / Non-finite screening magnitude cap
END_VAR

(* —— 段 1：输出缺省与样本数闸（纯函数，每调用重算） —— *)
fK1 := 0.0;  fK2 := 0.0;  fB := 0.0;  fR2 := 0.0;      // 输出缺省全 0（不给看似可信数字）
bIdentifiable := FALSE;                                  // 缺省不可辨识（安全侧）
bDegenerate   := FALSE;                                  // 缺省未退化
nErrId := 16#0000_0000;                                  // 事件码缺省无事件
FC_DL_LinearRegression2Var := FALSE;                     // 返回值缺省失败

IF (nSampleCount < 4) OR (nSampleCount > nMaxSmp) THEN
    nErrId := 16#0005_0202;                              // 故障级：样本不足或超数组上界
    RETURN;                                                // 不进入求解
END_IF

(* —— 段 2：累加矩 + 非有限值整批筛查（NaN 用 x<>x 自反判定，Inf 用幅值上限兜） —— *)
rN := LREAL(nSampleCount);
FOR k := 0 TO (nSampleCount - 1) DO
    bFin := (afX1[k] = afX1[k]) AND (afX2[k] = afX2[k]) AND (afY[k] = afY[k])
            AND (ABS(afX1[k]) < rFinLim) AND (ABS(afX2[k]) < rFinLim) AND (ABS(afY[k]) < rFinLim);
    IF NOT bFin THEN
        nErrId := 16#0005_0302;                          // 故障级：样本含非有限值，整批无效
        RETURN;                                            // 不污染统计
    END_IF
    rDx1 := LREAL(afX1[k]);  rDx2 := LREAL(afX2[k]);  rDy := LREAL(afY[k]);
    rSx1 := rSx1 + rDx1;  rSx2 := rSx2 + rDx2;  rSy := rSy + rDy;
    rS11 := rS11 + rDx1 * rDx1;  rS22 := rS22 + rDx2 * rDx2;
    rS12 := rS12 + rDx1 * rDx2;  rS1y := rS1y + rDx1 * rDy;  rS2y := rS2y + rDx2 * rDy;
    rSyy := rSyy + rDy * rDy;
END_FOR

(* —— 段 3：中心化方差/协方差与共线性判据 —— *)
rM1 := rSx1 / rN;  rM2 := rSx2 / rN;  rMy := rSy / rN;   // 均值（rN >= 4，无除零）
rV1 := rS11 - rSx1 * rM1;  rV2 := rS22 - rSx2 * rM2;  rC12 := rS12 - rSx1 * rM2;
IF (rV1 < rDetFloor) OR (rV2 < rDetFloor) THEN
    bDegenerate := TRUE;                                  // x1 或 x2 无离散：正规方程退化
    nErrId := 16#0005_0402;                               // 故障级：退化
    RETURN;
END_IF
rR12 := rC12 / SQRT(rV1 * rV2);                           // 相关系数（分母已闸）
IF ABS(rR12) > LREAL(fCollinearLimit) THEN
    nErrId := 16#0005_0102;                               // 信息级：共线性越限，判不可辨识
    bIdentifiable := FALSE;                               // 不输出斜率（防病态解误导）
    FC_DL_LinearRegression2Var := TRUE;                   // 求解已执行但结果判不可辨识
    RETURN;
END_IF

(* —— 段 4：3x3 正规方程 Cramer 求解（|det| < 1E-12 判退化） —— *)
rDet := rN * (rS11 * rS22 - rS12 * rS12)
      - rSx1 * (rSx1 * rS22 - rS12 * rSx2)
      + rSx2 * (rSx1 * rS12 - rS11 * rSx2);               // 3x3 行列式
IF ABS(rDet) < rDetFloor THEN
    bDegenerate := TRUE;                                  // 退化标志
    nErrId := 16#0005_0402;                               // 故障级：正规方程退化
    RETURN;
END_IF
fB  := REAL((rSy  * (rS11 * rS22 - rS12 * rS12)
           - rSx1 * (rS1y * rS22 - rS12 * rS2y)
           + rSx2 * (rS1y * rS12 - rS11 * rS2y)) / rDet); // 截距 b（第一列替换为 RHS 的行列式）
fK1 := REAL((rN   * (rS1y * rS22 - rS12 * rS2y)
           - rSy  * (rSx1 * rS22 - rS12 * rSx2)
           + rSx2 * (rSx1 * rS2y - rS1y * rSx2)) / rDet); // 斜率 k1（第二列替换为 RHS 的行列式）
fK2 := REAL((rN   * (rS11 * rS2y - rS1y * rS12)
           - rSx1 * (rSx1 * rS2y - rS1y * rSx2)
           + rSy  * (rSx1 * rS12 - rS11 * rSx2)) / rDet); // 斜率 k2（第三列替换为 RHS 的行列式）

(* —— 段 5：拟合优度 R²（SStot 近零防除零） —— *)
rSsTot := rSyy - rN * rMy * rMy;                          // 总平方和
IF rSsTot < rSsFloor THEN
    fR2 := 0.0;                                           // y 全等：R² 无定义，置 0 不给可信假象
    nErrId := 16#0005_0502;                               // 信息级：SStot 近零
ELSE
    rSsRes := 0.0;
    FOR k := 0 TO (nSampleCount - 1) DO
        rYhat := LREAL(fB) + LREAL(fK1) * LREAL(afX1[k]) + LREAL(fK2) * LREAL(afX2[k]);
        rSsRes := rSsRes + (LREAL(afY[k]) - rYhat) * (LREAL(afY[k]) - rYhat);
    END_FOR
    rDen := rSsTot;                                       // 分母已闸 > 1E-12
    fR2 := REAL(MAX(0.0, MIN(1.0, 1.0 - rSsRes / rDen))); // 钳到 0..1
END_IF

(* —— 段 6：出口标志与返回值 —— *)
bIdentifiable := TRUE;                                    // 走到此 = 共线性未越限且未退化
FC_DL_LinearRegression2Var := TRUE;                       // 求解成功

END_FUNCTION
